(* IEC 61131-3 sources: PLC-IsaVODE/PLC-IsaVODE/samples/plc-programs (part 15) *)

(* ---- 331-SCALE_B2.ST ---- *)
FUNCTION _BYTE_TO_REAL:REAL
	VAR_INPUT
		IN :	BYTE;
	END_VAR

	_BYTE_TO_REAL := USINT_TO_REAL(BYTE_TO_USINT(IN));
END_FUNCTION

FUNCTION SCALE_B2:REAL
	VAR_INPUT
		IN1 :	BYTE;
		IN2 :	BYTE;
		K :	REAL;
		O :	REAL;
		IN1_MIN :	REAL;
		IN1_MAX :	REAL;
		IN2_MIN :	REAL;
		IN2_MAX :	REAL;
	END_VAR

	SCALE_B2 := 	(((in1_max - in1_min)* _BYTE_TO_REAL(in1) + (in2_max - in2_min)* _BYTE_TO_REAL(in2)) * 0.003921569 + in1_min + in2_min) * K + O;

END_FUNCTION

PROGRAM program0
  VAR
	IN1 :	BYTE;
	IN2 :	BYTE;
	K :	REAL;
	O :	REAL;
	IN1_MIN :	REAL;
	IN1_MAX :	REAL;
	IN2_MIN :	REAL;
	IN2_MAX :	REAL;
	CEIL5_OUT : REAL;
  END_VAR

  CEIL5_OUT := SCALE_B2(IN1, IN2, K, O, IN1_MIN, IN1_MAX, IN2_MIN, IN2_MAX);

END_PROGRAM

CONFIGURATION Config0

  RESOURCE Res0 ON PLC
    TASK task0(INTERVAL := T#20ms,PRIORITY := 0);
    PROGRAM instance0 WITH task0 : program0;
  END_RESOURCE
END_CONFIGURATION

(* ---- 334-AIR_ENTHALPY.ST ---- *)
FUNCTION SDD:REAL

	VAR_INPUT
		T :	REAL;
		ICE :	BOOL;
	END_VAR

	IF ice THEN
		SDD := 611.153 * EXP(22.4433 * T / (272.186 + T));
	ELSE
		SDD := 611.213 * EXP(17.5043 * T / (241.2 + T));
	END_IF;

END_FUNCTION

FUNCTION DEW_CON:REAL

	VAR_INPUT
		RH :	REAL;
		T :	REAL;
	END_VAR

	IF RH > 0.0 AND T > -50.0 THEN
		DEW_CON := 2.166824303E-2 * RH * SDD(T,FALSE)  / (T - -273.15);
	ELSE
		DEW_CON := 0.0;
	END_IF;

END_FUNCTION

FUNCTION AIR_ENTHALPY:REAL

	VAR_INPUT
		T :	REAL;
		RH :	REAL;
	END_VAR

	Air_enthalpy := 1.00482 * T + (1.86 * T + 2500.78) * dew_con(RH,T);

END_FUNCTION

PROGRAM program0
  VAR
    T :	REAL;
	RH :	REAL;
    CEIL5_OUT : REAL;
  END_VAR

  CEIL5_OUT := AIR_ENTHALPY(T, RH);
END_PROGRAM

CONFIGURATION Config0

  RESOURCE Res0 ON PLC
    TASK task0(INTERVAL := T#20ms,PRIORITY := 0);
    PROGRAM instance0 WITH task0 : program0;
  END_RESOURCE
END_CONFIGURATION

(* ---- 335-FRMP_B.ST ---- *)
FUNCTION FRMP_B:BYTE

	VAR_INPUT
		START :	BYTE;
		DIR :	BOOL;
		TD :	TIME;
		TR :	TIME;
	END_VAR

	IF TD < TR THEN
		FRMP_B := MIN(UDINT_TO_BYTE(DWORD_TO_UDINT(SHL(TIME_TO_DWORD(TD), 8)) / TIME_TO_UDINT(TR)), SEL(DIR, START, USINT_TO_BYTE(USINT#255 - BYTE_TO_USINT(START))));
		IF DIR THEN
			FRMP_B := USINT_TO_BYTE(BYTE_TO_USINT(START) + BYTE_TO_USINT(FRMP_B));
		ELSE
			FRMP_B := USINT_TO_BYTE(BYTE_TO_USINT(START) - BYTE_TO_USINT(FRMP_B));
		END_IF;
	ELSE
		FRMP_B := SEL(DIR, BYTE#0, BYTE#255);
	END_IF;
END_FUNCTION

PROGRAM program0
  VAR
    LocalVar0 : BYTE;
	LocalVar1 : BOOL;
	LocalVar2 : TIME;
	LocalVar3 : TIME;
    LocalOUT  : BYTE;
  END_VAR

  LocalOUT := FRMP_B(LocalVar0, LocalVar1, LocalVar2,LocalVar3);
END_PROGRAM

CONFIGURATION Config0
  RESOURCE Res0 ON PLC
    TASK task0(INTERVAL := T#20ms,PRIORITY := 0);
    PROGRAM instance0 WITH task0 : program0;
  END_RESOURCE
END_CONFIGURATION

(* ---- 336-MD5_AUX.ST ---- *)
FUNCTION MD5_AUX:DWORD

	VAR_INPUT
		N :	INT;
		A :	DWORD;
		B :	DWORD;
		C :	DWORD;
		D :	DWORD;
		X :	DWORD;
		U :	INT;
		T :	DWORD;
	END_VAR

	VAR
		w :	DWORD;
	END_VAR

	CASE N OF
		1: w := (B AND C) OR (NOT(B) AND D);
		2: w := (B AND D) OR (C AND NOT D);
		3: w := (B XOR C XOR D);
		4: w := (C XOR (B OR  NOT(D)));
	END_CASE;

	MD5_AUX := UDINT_TO_DWORD(DWORD_TO_UDINT(B) + DWORD_TO_UDINT(ROL_DWORD(UDINT_TO_DWORD(DWORD_TO_UDINT(A) + DWORD_TO_UDINT(w) + DWORD_TO_UDINT(X) + DWORD_TO_UDINT(T)),U)));

END_FUNCTION

PROGRAM program0
	VAR
		N :	INT;
		A :	DWORD;
		B :	DWORD;
		C :	DWORD;
		D :	DWORD;
		X :	DWORD;
		U :	INT;
		T :	DWORD;
		CEIL5_OUT : DWORD;
	END_VAR

  	CEIL5_OUT := MD5_AUX(N, A, B, C, D, X, U, T);
END_PROGRAM

CONFIGURATION Config0

  RESOURCE Res0 ON PLC
    TASK task0(INTERVAL := T#20ms,PRIORITY := 0);
    PROGRAM instance0 WITH task0 : program0;
  END_RESOURCE
END_CONFIGURATION

(* ---- 34-TIME_TO_INT.ST ---- *)
FUNCTION TIME_TO_INT1:INT

VAR_INPUT
	IN :	TIME;
END_VAR

TIME_TO_INT1 := DINT_TO_INT(TIME_TO_DINT(IN));
END_FUNCTION

PROGRAM program0
  VAR
	IN :	TIME;
    CEIL5_OUT : INT;
  END_VAR

  CEIL5_OUT := TIME_TO_INT1(IN);
END_PROGRAM

CONFIGURATION Config0

  RESOURCE Res0 ON PLC
    TASK task0(INTERVAL := T#20ms,PRIORITY := 0);
    PROGRAM instance0 WITH task0 : program0;
  END_RESOURCE
END_CONFIGURATION

(* ---- 35-C_TO_F.ST ---- *)
FUNCTION C_TO_F:REAL
	VAR_INPUT
		CELSIUS :	REAL;
	END_VAR

	C_TO_F := celsius * 1.8 + 32.0;
END_FUNCTION

PROGRAM program0
  VAR
    LocalVar0 : REAL;
    CEIL5_OUT : REAL;
  END_VAR

  CEIL5_OUT := C_TO_F(LocalVar0);
END_PROGRAM

CONFIGURATION Config0

  RESOURCE Res0 ON PLC
    TASK task0(INTERVAL := T#20ms,PRIORITY := 0);
    PROGRAM instance0 WITH task0 : program0;
  END_RESOURCE
END_CONFIGURATION

(* ---- 355-MULTIME.ST ---- *)
FUNCTION _REAL_TO_DWORD: DWORD

  VAR_INPUT
    X :	REAL;
  END_VAR

  IF REAL_TO_DWORD(0.5) = DWORD#1 THEN
    _REAL_TO_DWORD := REAL_TO_DWORD(x);
  ELSIF X > 0.0 THEN
    _REAL_TO_DWORD := REAL_TO_DWORD(x+0.5);
  ELSIF X < 0.0 THEN
    _REAL_TO_DWORD := REAL_TO_DWORD(x-0.5);
  ELSE
    _REAL_TO_DWORD := DWORD#0;
  END_IF;
END_FUNCTION

FUNCTION _DWORD_TO_REAL:REAL
	VAR_INPUT
		IN :	DWORD;
	END_VAR

	_DWORD_TO_REAL := UDINT_TO_REAL(DWORD_TO_UDINT(IN));

END_FUNCTION

FUNCTION MULTIME:TIME
	VAR_INPUT
		T :	TIME;
		M :	REAL;
	END_VAR

	multime := DWORD_TO_TIME(_REAL_TO_DWORD(_DWORD_TO_REAL(TIME_TO_DWORD(t))*M));
END_FUNCTION

PROGRAM program0
  VAR
    LocalVar0 : TIME;
	LocalVar1 : REAL;
	LocalOUT  : TIME;
  END_VAR
  	LocalOUT := MULTIME(LocalVar0, LocalVar1);
END_PROGRAM

CONFIGURATION Config0
  RESOURCE Res0 ON PLC
    TASK task0(INTERVAL := T#20ms,PRIORITY := 0);
    PROGRAM instance0 WITH task0 : program0;
  END_RESOURCE
END_CONFIGURATION

(* ---- 356-OFFSET2.ST ---- *)
FUNCTION OFFSET2:REAL

	VAR_INPUT
		X :	REAL;
		O1 :	BOOL;
		O2 :	BOOL;
		O3 :	BOOL;
		O4 :	BOOL;
		D :	BOOL;
		OFFSET_1 :	REAL;
		OFFSET_2 :	REAL;
		OFFSET_3 :	REAL;
		OFFSET_4 :	REAL;
		DEFAULT :	REAL;
	END_VAR

	IF D THEN Offset2 := default; ELSE Offset2 := X; END_IF;
	IF O4 THEN Offset2 := Offset2 + offset_4;
	ELSIF O3 THEN Offset2 := Offset2 + offset_3;
	ELSIF O2 THEN Offset2 := Offset2 + offset_2;
	ELSIF O1 THEN Offset2 := Offset2 + offset_1;
	END_IF;

END_FUNCTION

PROGRAM program0
	VAR
		X :	REAL;
		O1 :	BOOL;
		O2 :	BOOL;
		O3 :	BOOL;
		O4 :	BOOL;
		D :	BOOL;
		OFFSET_1 :	REAL;
		OFFSET_2 :	REAL;
		OFFSET_3 :	REAL;
		OFFSET_4 :	REAL;
		DEFAULT :	REAL;
		OUT : REAL;
	END_VAR

	OUT := OFFSET2(X, O1, O2, O3, O4, D, OFFSET_1, OFFSET_2, OFFSET_3, OFFSET_4, DEFAULT);
END_PROGRAM

CONFIGURATION Config0

	RESOURCE Res0 ON PLC
		TASK task0(INTERVAL := T#20ms,PRIORITY := 0);
		PROGRAM instance0 WITH task0 : program0;
	END_RESOURCE

END_CONFIGURATION

(* ---- 36-DATE_TO_UDINT.ST ---- *)
FUNCTION DATE_TO_UDINT2:UDINT
	VAR_INPUT
		IN :	UDINT;
	END_VAR

	DATE_TO_UDINT2 := IN;
END_FUNCTION

PROGRAM program0
  VAR
    LocalVar0 : UDINT;
	LocalOUT  : UDINT;
  END_VAR
  	LocalOUT := DATE_TO_UDINT2(LocalVar0);
END_PROGRAM

CONFIGURATION Config0
  RESOURCE Res0 ON PLC
    TASK task0(INTERVAL := T#20ms,PRIORITY := 0);
    PROGRAM instance0 WITH task0 : program0;
  END_RESOURCE
END_CONFIGURATION

(* ---- 363-OFFSET.ST ---- *)
FUNCTION _OFFSET:REAL

	VAR_INPUT
		X :	REAL;
		O1 :	BOOL;
		O2 :	BOOL;
		O3 :	BOOL;
		O4 :	BOOL;
		D :	BOOL;
		OFFSET_1 :	REAL;
		OFFSET_2 :	REAL;
		OFFSET_3 :	REAL;
		OFFSET_4 :	REAL;
		DEFAULT :	REAL;
	END_VAR

	IF D THEN _Offset := default; ELSE _Offset := X; END_IF;
	IF O1 THEN _Offset := _Offset + offset_1; END_IF;
	IF O2 THEN _Offset := _Offset + offset_2; END_IF;
	IF O3 THEN _Offset := _Offset + offset_3; END_IF;
	IF O4 THEN _Offset := _Offset + offset_4; END_IF;

END_FUNCTION

PROGRAM program0

	VAR
		X :	REAL;
		O1 :	BOOL;
		O2 :	BOOL;
		O3 :	BOOL;
		O4 :	BOOL;
		D :	BOOL;
		OFFSET_1 :	REAL;
		OFFSET_2 :	REAL;
		OFFSET_3 :	REAL;
		OFFSET_4 :	REAL;
		DEFAULT :	REAL;
		OUT : REAL;
	END_VAR

	OUT := _OFFSET(X, O1, O2, O3, O4, D, OFFSET_1, OFFSET_2, OFFSET_3, OFFSET_4, DEFAULT);
END_PROGRAM

CONFIGURATION Config0

	RESOURCE Res0 ON PLC
		TASK task0(INTERVAL := T#20ms,PRIORITY := 0);
		PROGRAM instance0 WITH task0 : program0;
	END_RESOURCE

END_CONFIGURATION

(* ---- 365-CMP.ST ---- *)
FUNCTION EXP10 : REAL
  VAR_INPUT
    x : REAL;
  END_VAR

  exp10 := EXP(X * 2.30258509299405);
  (* from OSCAT library; www.oscat.de  *)
END_FUNCTION

FUNCTION FLOOR : INT
  VAR_INPUT
    x : REAL;
  END_VAR

  FLOOR := REAL_TO_INT(X);
  IF INT_TO_REAL(FLOOR) > X THEN
  	floor := floor - 1;
  END_IF;
  (* from OSCAT library; www.oscat.de  *)
END_FUNCTION

FUNCTION CMP:BOOL
	VAR_INPUT
		X :	REAL;
		Y :	REAL;
		N :	INT;
	END_VAR

	VAR
		tmp :	REAL;
	END_VAR

	tmp := ABS(x);
	IF tmp > 0.0 THEN
		tmp := EXP10(INT_TO_REAL(FLOOR(LOG(tmp))-N+1));
	ELSE
		tmp := EXP10(tmp);
	END_IF;
	CMP := ABS(X - Y) < tmp;

END_FUNCTION

PROGRAM program0
  VAR
    LocalVar0 : REAL;
    LocalVar1 : REAL;
	LocalVar2 : INT;
    CEIL5_OUT : BOOL;
  END_VAR

  CEIL5_OUT := CMP(LocalVar0, LocalVar1, LocalVar2);
END_PROGRAM

CONFIGURATION Config0

  RESOURCE Res0 ON PLC
    TASK task0(INTERVAL := T#20ms,PRIORITY := 0);
    PROGRAM instance0 WITH task0 : program0;
  END_RESOURCE
END_CONFIGURATION

(* ---- 37-LEAP_DAY.ST ---- *)
FUNCTION LEAP_DAY:BOOL

	VAR_INPUT
		IDATE :	UDINT;
	END_VAR

	LEAP_DAY := IDATE MOD UDINT#126230400 = UDINT#68169600;

END_FUNCTION

PROGRAM program0
	VAR
		IDATE :	UDINT;
		OUT : BOOL;
	END_VAR

	OUT := LEAP_DAY(IDATE);
END_PROGRAM

CONFIGURATION Config0

	RESOURCE Res0 ON PLC
		TASK task0(INTERVAL := T#20ms,PRIORITY := 0);
		PROGRAM instance0 WITH task0 : program0;
	END_RESOURCE

END_CONFIGURATION

(* ---- 370-SET_TOD.ST ---- *)
FUNCTION _REAL_TO_UDINT:UDINT

	VAR_INPUT
		X :	REAL;
	END_VAR

	IF REAL_TO_UDINT(0.5) = UDINT#1 THEN
		_REAL_TO_UDINT := REAL_TO_UDINT(x);
	ELSIF X > 0.0 THEN
		_REAL_TO_UDINT := REAL_TO_UDINT(x+0.5);
	ELSIF X < 0.0 THEN
		_REAL_TO_UDINT := REAL_TO_UDINT(x-0.5);
	ELSE
		_REAL_TO_UDINT := UDINT#0;
	END_IF;

END_FUNCTION

FUNCTION _INT_TO_UDINT:UDINT

	VAR_INPUT
		IN :	INT;
	END_VAR

	_INT_TO_UDINT := DINT_TO_UDINT(INT_TO_DINT(IN));

END_FUNCTION

FUNCTION SET_TOD:UDINT

	VAR_INPUT
		HOUR :	INT;
		MINUTE :	INT;
		SECOND :	REAL;
	END_VAR

	set_Tod := _REAL_TO_UDINT(second * 1000.0) + _INT_TO_UDINT(minute) * UDINT#60000 + _INT_TO_UDINT(hour) * UDINT#3600000;

END_FUNCTION

PROGRAM program0

	VAR
		HOUR :	INT;
		MINUTE :	INT;
		SECOND :	REAL;
		CEIL5_OUT : UDINT;
	END_VAR

	CEIL5_OUT := SET_TOD(HOUR, MINUTE, SECOND);

END_PROGRAM

CONFIGURATION Config0

	RESOURCE Res0 ON PLC
		TASK task0(INTERVAL := T#20ms,PRIORITY := 0);
		PROGRAM instance0 WITH task0 : program0;
	END_RESOURCE

END_CONFIGURATION

(* ---- 371-HEAT_INDEX.ST ---- *)
FUNCTION C_TO_F:REAL
	VAR_INPUT
		CELSIUS :	REAL;
	END_VAR

	C_TO_F := celsius * 1.8 + 32.0;
END_FUNCTION

FUNCTION F_TO_C:REAL
	VAR_INPUT
		FAHRENHEIT :	REAL;
	END_VAR
	F_TO_C := (fahrenheit - 32.0) * 0.5555555555555;
END_FUNCTION

FUNCTION HEAT_INDEX:REAL

	VAR_INPUT
		T :	REAL;
		RH :	REAL;
	END_VAR

	VAR
		RH2 :	REAL;
		T2 :	REAL;
		TX :	REAL;
	END_VAR

	IF RH < 20.0 OR T < 20.0 THEN
		HEAT_INDEX := T;
	ELSE
		TX := T;
		RH2 := RH * RH;
		TX := C_TO_F(TX);
		T2 := TX * TX;
		HEAT_INDEX := -42.379 + 2.04901523 * TX - 6.83783E-3 * T2
				+ RH * (10.1433127 - 0.22475541 * TX + 1.22874E-3 * T2)
				+ RH2 * (8.5282E-4 * TX - 5.481717E-2 - 1.99E-6 * T2);
		HEAT_INDEX := F_TO_C(HEAT_INDEX);
	END_IF;

END_FUNCTION

PROGRAM program0
  VAR
    T :	REAL;
	RH :	REAL;
    CEIL5_OUT : REAL;
  END_VAR

  CEIL5_OUT := HEAT_INDEX(T, RH);
END_PROGRAM

CONFIGURATION Config0

  RESOURCE Res0 ON PLC
    TASK task0(INTERVAL := T#20ms,PRIORITY := 0);
    PROGRAM instance0 WITH task0 : program0;
  END_RESOURCE
END_CONFIGURATION

(* ---- 38-TOD_TO_TIME.ST ---- *)
FUNCTION TOD_TO_TIME:TIME
	VAR_INPUT
		IN :	UDINT;
	END_VAR

	TOD_TO_TIME := DWORD_TO_TIME(UDINT_TO_DWORD(IN));
END_FUNCTION

PROGRAM program0
  VAR
	IN :	UDINT;
    CEIL5_OUT : TIME;
  END_VAR

  CEIL5_OUT := TOD_TO_TIME(IN);
END_PROGRAM

CONFIGURATION Config0

  RESOURCE Res0 ON PLC
    TASK task0(INTERVAL := T#20ms,PRIORITY := 0);
    PROGRAM instance0 WITH task0 : program0;
  END_RESOURCE
END_CONFIGURATION

(* ---- 384-EXPN.ST ---- *)
FUNCTION BIT_OF_DWORD : BOOL
  VAR_INPUT
    IN : DWORD;
    N : INT;
  END_VAR

  BIT_OF_DWORD := (SHR(in,N) AND 16#00000001) > 0;
END_FUNCTION

FUNCTION EXPN:REAL

	VAR_INPUT
		X :	REAL;
		N :	INT;
	END_VAR

	VAR
		N_word :	WORD;
		X_tmp :	REAL;
		sign :	BOOL;
	END_VAR

	N_word := INT_TO_WORD(N);
	X_tmp := X;
	sign := BIT_OF_DWORD(WORD_TO_DWORD(N_word),15);
	N_word := INT_TO_WORD(ABS(N));
	IF BIT_OF_DWORD(WORD_TO_DWORD(N_word),0) THEN expn := X_tmp; ELSE expn := 1.0; END_IF;    (* N_word.X0 *)
	N_word := SHR(N_word,1);
	WHILE N_word > WORD#0 DO
		X_tmp := X_tmp * X_tmp;
		IF BIT_OF_DWORD(WORD_TO_DWORD(N_word),0) THEN expn := expn * X_tmp; END_IF;       (* N_word.X0 *)
		N_word := SHR(N_word,1);
	END_WHILE;
	IF sign THEN EXPN := 1.0 / EXPN; END_IF;

END_FUNCTION

PROGRAM program0
  VAR
    LocalVar0 : REAL;
	LocalVar1 : INT;
	LocalOUT  : REAL;
  END_VAR
  	LocalOUT := EXPN(LocalVar0, LocalVar1);
END_PROGRAM

CONFIGURATION Config0
  RESOURCE Res0 ON PLC
    TASK task0(INTERVAL := T#20ms,PRIORITY := 0);
    PROGRAM instance0 WITH task0 : program0;
  END_RESOURCE
END_CONFIGURATION

(* ---- 385-ROUND.ST ---- *)
FUNCTION _REAL_TO_DINT:DINT
	VAR_INPUT
		X :	REAL;
	END_VAR

	IF REAL_TO_DINT(0.5) = DINT#1 THEN
		_REAL_TO_DINT := REAL_TO_DINT(x);
		RETURN;
	END_IF;

	IF X > 0.0 THEN
		_REAL_TO_DINT := REAL_TO_DINT(x+0.5);
	ELSIF X < 0.0 THEN
		_REAL_TO_DINT := REAL_TO_DINT(x-0.5);
	ELSE
		_REAL_TO_DINT := DINT#0;
	END_IF;
END_FUNCTION

FUNCTION ROUND:REAL

	VAR_INPUT
		IN :	REAL;
		N :	INT;
	END_VAR

	VAR
		X :	REAL;
	END_VAR

	IF N < 4 THEN
		IF N < 2 THEN
			IF N = 0 THEN X := 1.0; ELSE X := 10.0; END_IF;
		ELSE
			IF N = 2 THEN X := 100.0; ELSE X := 1000.0; END_IF;
		END_IF;
	ELSE
		IF N < 6 THEN
			IF N = 4 THEN X := 10000.0; ELSE X := 100000.0; END_IF;
		ELSE
			IF N = 6 THEN X := 1000000.0; ELSE X := 10000000.0; END_IF;
		END_IF;
	END_IF;

	ROUND := DINT_TO_REAL(_REAL_TO_DINT(in * X)) / X;

END_FUNCTION

PROGRAM program0
	VAR
		IN : REAL;
		N :	INT;
		X :	REAL;
	END_VAR
		X := ROUND(IN, N);
END_PROGRAM

CONFIGURATION Config0

	RESOURCE Res0 ON PLC
		TASK task0(INTERVAL := T#20ms,PRIORITY := 0);
		PROGRAM instance0 WITH task0 : program0;
	END_RESOURCE

END_CONFIGURATION

(* ---- 39-DATE_TO_REAL.ST ---- *)
FUNCTION DATE_TO_REAL2:REAL
	VAR_INPUT
		IN :	UDINT;
	END_VAR

	DATE_TO_REAL2 := UDINT_TO_REAL(IN);
END_FUNCTION

PROGRAM program0
  VAR
    LocalVar0 : UDINT;
	LocalOUT  : REAL;
  END_VAR
  	LocalOUT := DATE_TO_REAL2(LocalVar0);
END_PROGRAM

CONFIGURATION Config0
  RESOURCE Res0 ON PLC
    TASK task0(INTERVAL := T#20ms,PRIORITY := 0);
    PROGRAM instance0 WITH task0 : program0;
  END_RESOURCE
END_CONFIGURATION

(* ---- 395-SET_DATE.ST ---- *)
FUNCTION _INT_TO_UDINT:UDINT
	VAR_INPUT
		IN :	INT;
	END_VAR

	_INT_TO_UDINT := DINT_TO_UDINT(INT_TO_DINT(IN));
END_FUNCTION

FUNCTION SET_DATE:UDINT

	VAR_INPUT
		YEAR :	INT;
		MONTH :	INT;
		DAY :	INT;
	END_VAR

	VAR
		count :	INT;
	END_VAR

	IF month > 2 THEN
		count := (month - 1) * 30;
		IF month > 7 THEN
			count := count + DWORD_TO_INT(SHR(DINT_TO_DWORD(INT_TO_DINT(month) - INT_TO_DINT(3)),1));
		ELSE
			count := count + DWORD_TO_INT(SHR(DINT_TO_DWORD(INT_TO_DINT(month) - INT_TO_DINT(4)),1));
		END_IF;
		IF SHL(INT_TO_WORD(year),14) = WORD#0 THEN
			count := count + 1;
		END_IF;
	ELSE
		count := (month - 1) * 31;
	END_IF;
	SET_DATE := (_INT_TO_UDINT(count + day - 1) + DWORD_TO_UDINT(SHR(UDINT_TO_DWORD(_INT_TO_UDINT(year) * UDINT#1461 - UDINT#2878169), 2))) * UDINT#86400;

END_FUNCTION

PROGRAM program0
  VAR
	YEAR :	INT;
	MONTH :	INT;
	DAY :	INT;
    CEIL5_OUT : UDINT;
  END_VAR

  CEIL5_OUT := SET_DATE(YEAR, MONTH, DAY);
END_PROGRAM

CONFIGURATION Config0

  RESOURCE Res0 ON PLC
    TASK task0(INTERVAL := T#20ms,PRIORITY := 0);
    PROGRAM instance0 WITH task0 : program0;
  END_RESOURCE
END_CONFIGURATION

(* ---- 40-DWORD_TO_DT.ST ---- *)
FUNCTION DWORD_TO_DT2:UDINT

	VAR_INPUT
		IN :	DWORD;
	END_VAR

	DWORD_TO_DT2 := DWORD_TO_UDINT(IN);
END_FUNCTION

PROGRAM program0
  VAR
    LocalVar0 : DWORD;
	LocalOUT  : UDINT;
  END_VAR
  	LocalOUT := DWORD_TO_DT2(LocalVar0);
END_PROGRAM

CONFIGURATION Config0
  RESOURCE Res0 ON PLC
    TASK task0(INTERVAL := T#20ms,PRIORITY := 0);
    PROGRAM instance0 WITH task0 : program0;
  END_RESOURCE
END_CONFIGURATION

(* ---- 400-TEMP_PT.ST ---- *)
FUNCTION RES_PT:REAL
	VAR_INPUT
		T :	REAL;
		R0 :	REAL;
	END_VAR

	VAR
		T2 :	REAL;
	END_VAR

	T2 := T * T;

	IF T >= 0.0 THEN
		RES_PT := R0 * ( 1.0 + 3.90802E-3 * T + -5.802E-7 * T2);
	ELSE
		RES_PT := R0 * ( 1.0 + 3.90802E-3 * T + -5.802E-7 * T2 + -4.27350E-12 * (T - 100.0) * T2 * T);
	END_IF;

END_FUNCTION

FUNCTION TEMP_PT:REAL

	VAR_INPUT
		RES :	REAL;
		R0 :	REAL;
	END_VAR

	VAR
		step_var :	REAL := REAL#50.0;
		X :	REAL;
		Y :	REAL;
		t1 :	REAL;
	END_VAR

	X := 3.9083E-3 * R0;
	Y := -5.775E-7 * R0;
	IF Res >= R0 THEN
		t1 := X * X - 4.0 * Y * (R0 - Res);
		IF t1 < 0.0 THEN
			TEMP_PT := 10000.0;
		ELSE
			TEMP_PT := (-X + SQRT(t1)) / (2.0 * Y);
		END_IF;
	ELSE
		TEMP_PT := -100.0;
		WHILE step_var > 0.01 DO
			IF RES_PT(TEMP_PT, R0) < res THEN TEMP_PT := TEMP_PT + step_var; ELSE TEMP_PT := TEMP_PT - step_var; END_IF;
			step_var := step_var * 0.5;
		END_WHILE;
	END_IF;
END_FUNCTION

PROGRAM program0
	VAR
		RES :	REAL;
		R0 :	REAL;
		CEIL5_OUT : REAL;
	END_VAR

	CEIL5_OUT := TEMP_PT(RES, R0);
END_PROGRAM

CONFIGURATION Config0
	RESOURCE Res0 ON PLC
		TASK task0(INTERVAL := T#20ms,PRIORITY := 0);
		PROGRAM instance0 WITH task0 : program0;
	END_RESOURCE
END_CONFIGURATION

(* ---- 404-MONTH_OF_DATE.ST ---- *)
FUNCTION LEAP_OF_DATE:BOOL

	VAR_INPUT
		IDATE :	UDINT;
	END_VAR

	LEAP_OF_DATE := SHL(UDINT_TO_DWORD((idate + UDINT#43200) / UDINT#31557600), 30) = DWORD#16#80000000;

END_FUNCTION

FUNCTION DAY_OF_YEAR:INT
	VAR_INPUT
		IDATE :	DATE;
	END_VAR

	DAY_OF_YEAR := UDINT_TO_INT((DATE_TO_UDINT(idate) / UDINT#86400) MOD UDINT#1461);
	IF DAY_OF_YEAR > 729 THEN
		IF DAY_OF_YEAR > 1095 THEN DAY_OF_YEAR := DAY_OF_YEAR - 1095; ELSE DAY_OF_YEAR := DAY_OF_YEAR - 729; END_IF;
	ELSIF DAY_OF_YEAR > 364 THEN
		DAY_OF_YEAR := DAY_OF_YEAR - 364;
	ELSE
		DAY_OF_YEAR := DAY_OF_YEAR + 1;
	END_IF;
END_FUNCTION

FUNCTION MONTH_OF_DATE:INT

	VAR_INPUT
		IDATE :	DATE;
	END_VAR

	MONTH_OF_DATE := DAY_OF_YEAR(idate);
	IF MONTH_OF_DATE < 32 THEN
		MONTH_OF_DATE := 1;
	ELSIF LEAP_OF_DATE(DATE_TO_UDINT(IDATE)) THEN
		MONTH_OF_DATE := (MONTH_OF_DATE * 53 + 1668) / 1623;
	ELSE
		MONTH_OF_DATE := (MONTH_OF_DATE * 53 + 1700) / 1620;
	END_IF;

END_FUNCTION

PROGRAM program0
  VAR
    LocalVar0 : DATE;
	LocalOUT  : INT;
  END_VAR
  	LocalOUT := MONTH_OF_DATE(LocalVar0);
END_PROGRAM

CONFIGURATION Config0
  RESOURCE Res0 ON PLC
    TASK task0(INTERVAL := T#20ms,PRIORITY := 0);
    PROGRAM instance0 WITH task0 : program0;
  END_RESOURCE
END_CONFIGURATION

(* ---- 405-SCALE_B4.ST ---- *)
FUNCTION _BYTE_TO_REAL:REAL
	VAR_INPUT
		IN :	BYTE;
	END_VAR

	_BYTE_TO_REAL := USINT_TO_REAL(BYTE_TO_USINT(IN));
END_FUNCTION

FUNCTION SCALE_B4:REAL

	VAR_INPUT
		IN1 :	BYTE;
		IN2 :	BYTE;
		IN3 :	BYTE;
		IN4 :	BYTE;
		K :	REAL;
		O :	REAL;
		IN1_MIN :	REAL;
		IN1_MAX :	REAL;
		IN2_MIN :	REAL;
		IN2_MAX :	REAL;
		IN3_MIN :	REAL;
		IN3_MAX :	REAL;
		IN4_MIN :	REAL;
		IN4_MAX :	REAL;
	END_VAR

	SCALE_B4 := 	(((in1_max - in1_min)* _BYTE_TO_REAL(in1) + (in2_max - in2_min)* _BYTE_TO_REAL(in2) + (in3_max - in3_min)* _BYTE_TO_REAL(in3) + (in4_max - in4_min)* _BYTE_TO_REAL(in4))* 0.003921569 + in1_min + in2_min + in3_min + in4_min) * K + O;

END_FUNCTION

PROGRAM program0
  VAR
	IN1 :	BYTE;
	IN2 :	BYTE;
	IN3 :	BYTE;
	IN4 :	BYTE;
	K :	REAL;
	O :	REAL;
	IN1_MIN :	REAL;
	IN1_MAX :	REAL;
	IN2_MIN :	REAL;
	IN2_MAX :	REAL;
	IN3_MIN :	REAL;
	IN3_MAX :	REAL;
	IN4_MIN :	REAL;
	IN4_MAX :	REAL;
	CEIL5_OUT : REAL;
  END_VAR

  CEIL5_OUT := SCALE_B4(IN1, IN2, IN3, IN4, K, O, IN1_MIN, IN1_MAX, IN2_MIN, IN2_MAX, IN3_MIN, IN3_MAX, IN4_MIN, IN4_MAX);

END_PROGRAM

CONFIGURATION Config0

  RESOURCE Res0 ON PLC
    TASK task0(INTERVAL := T#20ms,PRIORITY := 0);
    PROGRAM instance0 WITH task0 : program0;
  END_RESOURCE
END_CONFIGURATION

(* ---- 408-SCALE_X4.ST ---- *)
FUNCTION SCALE_X4:REAL
	VAR_INPUT
		IN1 :	BOOL;
		IN2 :	BOOL;
		IN3 :	BOOL;
		IN4 :	BOOL;
		K :	REAL;
		O :	REAL;
		IN1_MIN :	REAL;
		IN1_MAX :	REAL;
		IN2_MIN :	REAL;
		IN2_MAX :	REAL;
		IN3_MIN :	REAL;
		IN3_MAX :	REAL;
		IN4_MIN :	REAL;
		IN4_MAX :	REAL;
	END_VAR
	IF NOT in1 THEN scale_X4 := in1_min; ELSE scale_X4 := in1_max; END_IF;
	IF NOT in2 THEN scale_x4 := scale_x4 + in2_min; ELSE scale_x4 := scale_x4 + in2_max; END_IF;
	IF NOT in3 THEN scale_x4 := scale_x4 + in3_min; ELSE scale_x4 := scale_x4 + in3_max; END_IF;
	IF NOT in4 THEN scale_x4 := scale_x4 + in4_min; ELSE scale_x4 := scale_x4 + in4_max; END_IF;
	scale_X4 := scale_X4 * k + O;
	END_FUNCTION

PROGRAM program0

  	VAR
		IN1 :	BOOL;
		IN2 :	BOOL;
		IN3 :	BOOL;
		IN4 :	BOOL;
		K :	REAL;
		O :	REAL;
		IN1_MIN :	REAL;
		IN1_MAX :	REAL;
		IN2_MIN :	REAL;
		IN2_MAX :	REAL;
		IN3_MIN :	REAL;
		IN3_MAX :	REAL;
		IN4_MIN :	REAL;
		IN4_MAX :	REAL;
		CEIL5_OUT : REAL;
  	END_VAR

  	CEIL5_OUT := SCALE_X4(IN1, IN2, IN3, IN4, K, O, IN1_MIN, IN1_MAX, IN2_MIN, IN2_MAX, IN3_MIN, IN3_MAX, IN4_MIN, IN4_MAX);
END_PROGRAM

CONFIGURATION Config0

	RESOURCE Res0 ON PLC
		TASK task0(INTERVAL := T#20ms,PRIORITY := 0);
		PROGRAM instance0 WITH task0 : program0;
	END_RESOURCE

END_CONFIGURATION

(* ---- 41-BYTE_TO_GRAY.ST ---- *)
FUNCTION BYTE_TO_GRAY:BYTE
	VAR_INPUT
		IN :	BYTE;
	END_VAR

	BYTE_TO_GRAY := IN XOR SHR(IN,1);
END_FUNCTION

PROGRAM program0
  VAR
    LocalVar0 : BYTE;
    CEIL5_OUT : BYTE;
  END_VAR

  CEIL5_OUT := BYTE_TO_GRAY(LocalVar0);
END_PROGRAM

CONFIGURATION Config0

  RESOURCE Res0 ON PLC
    TASK task0(INTERVAL := T#20ms,PRIORITY := 0);
    PROGRAM instance0 WITH task0 : program0;
  END_RESOURCE
END_CONFIGURATION

(* ---- 413-OSCAT_VERSION.ST ---- *)
FUNCTION _INT_TO_UDINT:UDINT
	VAR_INPUT
		IN :	INT;
	END_VAR

	_INT_TO_UDINT := DINT_TO_UDINT(INT_TO_DINT(IN));
END_FUNCTION

FUNCTION SET_DATE:UDINT

	VAR_INPUT
		YEAR :	INT;
		MONTH :	INT;
		DAY :	INT;
	END_VAR

	VAR
		count :	INT;
	END_VAR

	IF month > 2 THEN
		count := (month - 1) * 30;
		IF month > 7 THEN
			count := count + DWORD_TO_INT(SHR(DINT_TO_DWORD(INT_TO_DINT(month) - INT_TO_DINT(3)),1));
		ELSE
			count := count + DWORD_TO_INT(SHR(DINT_TO_DWORD(INT_TO_DINT(month) - INT_TO_DINT(4)),1));
		END_IF;
		IF SHL(INT_TO_WORD(year),14) = WORD#0 THEN
			count := count + 1;
		END_IF;
	ELSE
		count := (month - 1) * 31;
	END_IF;
	SET_DATE := (_INT_TO_UDINT(count + day - 1) + DWORD_TO_UDINT(SHR(UDINT_TO_DWORD(_INT_TO_UDINT(year) * UDINT#1461 - UDINT#2878169), 2))) * UDINT#86400;

END_FUNCTION

FUNCTION OSCAT_VERSION:DWORD

	VAR_INPUT
		IN :	BOOL;
	END_VAR

	IF in THEN
		Oscat_version := UDINT_TO_DWORD(set_Date(2012,01,02));
	ELSE
		Oscat_version := DWORD#333;
	END_IF;

END_FUNCTION

PROGRAM program0
	VAR
		IN :	BOOL;
		OUT : DWORD;
	END_VAR

	OUT := OSCAT_VERSION(IN);
END_PROGRAM

CONFIGURATION Config0

	RESOURCE Res0 ON PLC
		TASK task0(INTERVAL := T#20ms,PRIORITY := 0);
		PROGRAM instance0 WITH task0 : program0;
	END_RESOURCE

END_CONFIGURATION

(* ---- 417-NETWORK_VERSION.ST ---- *)
FUNCTION _INT_TO_UDINT:UDINT
	VAR_INPUT
		IN :	INT;
	END_VAR

	_INT_TO_UDINT := DINT_TO_UDINT(INT_TO_DINT(IN));
END_FUNCTION

FUNCTION SET_DATE:UDINT

	VAR_INPUT
		YEAR :	INT;
		MONTH :	INT;
		DAY :	INT;
	END_VAR

	VAR
		count :	INT;
	END_VAR

	IF month > 2 THEN
		count := (month - 1) * 30;
		IF month > 7 THEN
			count := count + DWORD_TO_INT(SHR(DINT_TO_DWORD(INT_TO_DINT(month) - INT_TO_DINT(3)),1));
		ELSE
			count := count + DWORD_TO_INT(SHR(DINT_TO_DWORD(INT_TO_DINT(month) - INT_TO_DINT(4)),1));
		END_IF;
		IF SHL(INT_TO_WORD(year),14) = WORD#0 THEN
			count := count + 1;
		END_IF;
	ELSE
		count := (month - 1) * 31;
	END_IF;
	SET_DATE := (_INT_TO_UDINT(count + day - 1) + DWORD_TO_UDINT(SHR(UDINT_TO_DWORD(_INT_TO_UDINT(year) * UDINT#1461 - UDINT#2878169), 2))) * UDINT#86400;

END_FUNCTION

FUNCTION NETWORK_VERSION:DWORD

	VAR_INPUT
		IN :	BOOL;
	END_VAR

	IF in THEN
		NETWORK_VERSION := UDINT_TO_DWORD(set_Date(2011,12,01));
	ELSE
		NETWORK_VERSION := DWORD#121;
	END_IF;

END_FUNCTION

PROGRAM program0
	VAR
		IN :	BOOL;
		CEIL5_OUT : DWORD;
	END_VAR

  	CEIL5_OUT := NETWORK_VERSION(IN);
END_PROGRAM

CONFIGURATION Config0

  RESOURCE Res0 ON PLC
    TASK task0(INTERVAL := T#20ms,PRIORITY := 0);
    PROGRAM instance0 WITH task0 : program0;
  END_RESOURCE
END_CONFIGURATION

(* ---- 419-BUILDING_VERSION.ST ---- *)
FUNCTION _INT_TO_UDINT:UDINT
	VAR_INPUT
		IN :	INT;
	END_VAR

	_INT_TO_UDINT := DINT_TO_UDINT(INT_TO_DINT(IN));
END_FUNCTION

FUNCTION SET_DATE:UDINT

	VAR_INPUT
		YEAR :	INT;
		MONTH :	INT;
		DAY :	INT;
	END_VAR

	VAR
		count :	INT;
	END_VAR

	IF month > 2 THEN
		count := (month - 1) * 30;
		IF month > 7 THEN
			count := count + DWORD_TO_INT(SHR(DINT_TO_DWORD(INT_TO_DINT(month) - INT_TO_DINT(3)),1));
		ELSE
			count := count + DWORD_TO_INT(SHR(DINT_TO_DWORD(INT_TO_DINT(month) - INT_TO_DINT(4)),1));
		END_IF;
		IF SHL(INT_TO_WORD(year),14) = WORD#0 THEN
			count := count + 1;
		END_IF;
	ELSE
		count := (month - 1) * 31;
	END_IF;
	SET_DATE := (_INT_TO_UDINT(count + day - 1) + DWORD_TO_UDINT(SHR(UDINT_TO_DWORD(_INT_TO_UDINT(year) * UDINT#1461 - UDINT#2878169), 2))) * UDINT#86400;

END_FUNCTION

FUNCTION BUILDING_VERSION:DWORD

	VAR_INPUT
		IN :	BOOL;
	END_VAR

	IF in THEN
		BUILDING_VERSION := UDINT_TO_DWORD(set_Date(2011,02,03));
	ELSE
		BUILDING_VERSION := DWORD#100;
	END_IF;

END_FUNCTION

PROGRAM program0
	VAR
		IN :	BOOL;
		CEIL5_OUT : DWORD;
	END_VAR

  	CEIL5_OUT := BUILDING_VERSION(IN);
END_PROGRAM

CONFIGURATION Config0

  RESOURCE Res0 ON PLC
    TASK task0(INTERVAL := T#20ms,PRIORITY := 0);
    PROGRAM instance0 WITH task0 : program0;
  END_RESOURCE
END_CONFIGURATION

(* ---- 42-F_TO_C.ST ---- *)
FUNCTION F_TO_C:REAL
	VAR_INPUT
		FAHRENHEIT :	REAL;
	END_VAR
	F_TO_C := (fahrenheit - 32.0) * 0.5555555555555;
END_FUNCTION

PROGRAM program0
  VAR
    LocalVar0 : REAL;
	LocalOUT  : REAL;
  END_VAR
  	LocalOUT := F_TO_C(LocalVar0);
END_PROGRAM

CONFIGURATION Config0
  RESOURCE Res0 ON PLC
    TASK task0(INTERVAL := T#20ms,PRIORITY := 0);
    PROGRAM instance0 WITH task0 : program0;
  END_RESOURCE
END_CONFIGURATION

(* ---- 421-GCD.ST ---- *)
FUNCTION GCD:INT

	VAR_INPUT
		A :	DINT;
		B :	DINT;
	END_VAR

	VAR
		t :	DINT;
		_A :	DINT;
		_B :	DINT;
	END_VAR

	_A := A;
	_B := B;

	IF _A = DINT#0 THEN
		GCD := DINT_TO_INT(ABS(_B));
	ELSIF _B = DINT#0 THEN
		GCD := DINT_TO_INT(ABS(_A));
	ELSE
		_A := ABS(_A);
		_B := ABS(_B);
		GCD := 1;

		WHILE NOT((DINT_TO_DWORD(_A) AND DWORD#1) > DWORD#0 OR (DINT_TO_DWORD(_B) AND DWORD#1) > DWORD#0) DO
			_A := DWORD_TO_DINT(SHR(DINT_TO_DWORD(_A),1));
			_B := DWORD_TO_DINT(SHR(DINT_TO_DWORD(_B),1));
			GCD := DWORD_TO_INT(SHR(INT_TO_DWORD(GCD),1));
		END_WHILE;
		WHILE _A > DINT#0 DO
			IF NOT((DINT_TO_DWORD(_A) AND DWORD#1) > DWORD#0) THEN
				_A := DWORD_TO_DINT(SHR(DINT_TO_DWORD(_A),1));
			ELSIF NOT((DINT_TO_DWORD(_B) AND DWORD#1) > DWORD#0) THEN
				_B := DWORD_TO_DINT(SHR(DINT_TO_DWORD(_B),1));
			ELSE
				t := DWORD_TO_DINT(SHR(DINT_TO_DWORD(ABS(_A-_B)),1));
				IF _A < _B THEN
					_B := t;
				ELSE
					_A := t;
				END_IF;
			END_IF;
		END_WHILE;
		GCD := GCD * DINT_TO_INT(_B);
	END_IF;

END_FUNCTION

PROGRAM program0
  VAR
    A :	DINT;
	B :	DINT;
    LocalOUT  : INT;
  END_VAR

  LocalOUT := GCD(A, B);
END_PROGRAM

CONFIGURATION Config0
  RESOURCE Res0 ON PLC
    TASK task0(INTERVAL := T#20ms,PRIORITY := 0);
    PROGRAM instance0 WITH task0 : program0;
  END_RESOURCE
END_CONFIGURATION

(* ---- 423-AIN.ST ---- *)
FUNCTION _BYTE_TO_INT:INT
	VAR_INPUT
		IN :	BYTE;
	END_VAR

	_BYTE_TO_INT := USINT_TO_INT(BYTE_TO_USINT(IN));
END_FUNCTION

FUNCTION _DWORD_TO_REAL:REAL
	VAR_INPUT
		IN :	DWORD;
	END_VAR

	_DWORD_TO_REAL := UDINT_TO_REAL(DWORD_TO_UDINT(IN));
END_FUNCTION

FUNCTION BIT_OF_DWORD:BOOL
	VAR_INPUT
		IN :	DWORD;
		N :	INT;
	END_VAR
	BIT_OF_DWORD := (SHR(in,n) AND DWORD#1) > DWORD#0;
END_FUNCTION

FUNCTION AIN:REAL
	VAR_INPUT
		IN :	DWORD;
		BITS :	BYTE;
		SIGN :	BYTE;
		LOW :	REAL;
		HIGH :	REAL;
	END_VAR

	VAR
		temp1 :	DWORD;
		temp2 :	DWORD;
		sx :	BOOL;
	END_VAR

	IF sign < BYTE#32 THEN
		temp1 := SHR(in, _BYTE_TO_INT(sign));
		sx := BIT_OF_DWORD(temp1,0); (* temp1.X0 *)
	ELSE
		sx := FALSE;
	END_IF;
	temp1 := SHR(DWORD#16#FFFFFFFF,32 - _BYTE_TO_INT(bits));
	temp2 := in AND temp1;
	AIN := (high - low)* _DWORD_TO_REAL(temp2) / _DWORD_TO_REAL(temp1) + low;
	IF sx THEN AIN := -AIN; END_IF;
END_FUNCTION

PROGRAM program0
  VAR
    LocalVar0 : DWORD;
	LocalVar1 : BYTE;
	LocalVar2 : BYTE;
	LocalVar3 : REAL;
	LocalVar4 : REAL;
    LocalOUT  : REAL;
  END_VAR

  LocalOUT := AIN(LocalVar0, LocalVar1, LocalVar2, LocalVar3, LocalVar4);
END_PROGRAM

CONFIGURATION Config0
  RESOURCE Res0 ON PLC
    TASK task0(INTERVAL := T#20ms,PRIORITY := 0);
    PROGRAM instance0 WITH task0 : program0;
  END_RESOURCE
END_CONFIGURATION

(* ---- 43-TANC.ST ---- *)
FUNCTION TANC:REAL

	VAR_INPUT
		X :	REAL;
	END_VAR

	IF X = 0.0 THEN
		TANC := 1.0;
	ELSE
		TANC := TAN(x) / x;
	END_IF;

END_FUNCTION

PROGRAM program0

	VAR
		X :	REAL;
		CEIL5_OUT : REAL;
	END_VAR

	CEIL5_OUT := TANC(X);

END_PROGRAM

CONFIGURATION Config0

	RESOURCE Res0 ON PLC
		TASK task0(INTERVAL := T#20ms,PRIORITY := 0);
		PROGRAM instance0 WITH task0 : program0;
	END_RESOURCE

END_CONFIGURATION

(* ---- 436-AOUT1.ST ---- *)
FUNCTION SIGN_R : BOOL
  VAR_INPUT
    IN : REAL;
  END_VAR

  SIGN_R := in < 0.0;
END_FUNCTION

FUNCTION _REAL_TO_DWORD: DWORD

  VAR_INPUT
    X :	REAL;
  END_VAR

  IF REAL_TO_DWORD(0.5) = DWORD#1 THEN
    _REAL_TO_DWORD := REAL_TO_DWORD(x);
  ELSIF X > 0.0 THEN
    _REAL_TO_DWORD := REAL_TO_DWORD(x+0.5);
  ELSIF X < 0.0 THEN
    _REAL_TO_DWORD := REAL_TO_DWORD(x-0.5);
  ELSE
    _REAL_TO_DWORD := DWORD#0;
  END_IF;
END_FUNCTION

FUNCTION AOUT1:DWORD

	VAR_INPUT
		IN :	REAL;
		BIT_0 :	INT;
		BIT_N :	INT;
		SIGN :	INT;
		LOW :	REAL;
		HIGH :	REAL;
	END_VAR

	VAR
		in2 :	REAL;
		sx :	BOOL;
	END_VAR

	IF sign < 32 THEN
		sx := sign_R(in);
		in2 := ABS(in);
	ELSE
		sx := FALSE;
		in2 := in;
	END_IF;

	in2 := LIMIT_REAL(low, in2, high);

	AOUT1 :=  SHL(_REAL_TO_DWORD((in2 - low) / (high - low) * UDINT_TO_REAL(DWORD_TO_UDINT(SHL(DWORD#2#1,bit_n - Bit_0 + 1)) - UDINT#1)),Bit_0);

	IF sx THEN AOUT1 := SHL(DWORD#2#1,sign) OR AOUT1; END_IF;

END_FUNCTION

PROGRAM program0
  VAR
    LocalVar0 : REAL;
	LocalVar1 : INT;
	LocalVar21 : INT;
	LocalVar2 : INT;
	LocalVar3 : REAL;
	LocalVar4 : REAL;
	LocalOUT  : DWORD;
  END_VAR
  	LocalOUT := AOUT1(LocalVar0, LocalVar1,LocalVar21, LocalVar2, LocalVar3,LocalVar4);
END_PROGRAM

CONFIGURATION Config0
  RESOURCE Res0 ON PLC
    TASK task0(INTERVAL := T#20ms,PRIORITY := 0);
    PROGRAM instance0 WITH task0 : program0;
  END_RESOURCE
END_CONFIGURATION

(* ---- 44-SETUP_EXTENDED_ASCII.ST ---- *)
FUNCTION SETUP_EXTENDED_ASCII:BOOL

	VAR_INPUT
		X :	BOOL;
	END_VAR

	SETUP_EXTENDED_ASCII := X OR TRUE;
END_FUNCTION

PROGRAM program0
  VAR
	X :	BOOL;
    CEIL5_OUT : BOOL;
  END_VAR

  CEIL5_OUT := SETUP_EXTENDED_ASCII(X);
END_PROGRAM

CONFIGURATION Config0

  RESOURCE Res0 ON PLC
    TASK task0(INTERVAL := T#20ms,PRIORITY := 0);
    PROGRAM instance0 WITH task0 : program0;
  END_RESOURCE
END_CONFIGURATION

(* ---- 443-SET_DT.ST ---- *)
FUNCTION _INT_TO_UDINT:UDINT
	VAR_INPUT
		IN :	INT;
	END_VAR

	_INT_TO_UDINT := DINT_TO_UDINT(INT_TO_DINT(IN));
END_FUNCTION

FUNCTION SET_DATE:UDINT

	VAR_INPUT
		YEAR :	INT;
		MONTH :	INT;
		DAY :	INT;
	END_VAR

	VAR
		count :	INT;
	END_VAR

	IF month > 2 THEN
		count := (month - 1) * 30;
		IF month > 7 THEN
			count := count + DWORD_TO_INT(SHR(DINT_TO_DWORD(INT_TO_DINT(month) - INT_TO_DINT(3)),1));
		ELSE
			count := count + DWORD_TO_INT(SHR(DINT_TO_DWORD(INT_TO_DINT(month) - INT_TO_DINT(4)),1));
		END_IF;
		IF SHL(INT_TO_WORD(year),14) = WORD#0 THEN
			count := count + 1;
		END_IF;
	ELSE
		count := (month - 1) * 31;
	END_IF;
	SET_DATE := (_INT_TO_UDINT(count + day - 1) + DWORD_TO_UDINT(SHR(UDINT_TO_DWORD(_INT_TO_UDINT(year) * UDINT#1461 - UDINT#2878169), 2))) * UDINT#86400;

END_FUNCTION

FUNCTION SET_DT:UDINT
	VAR_INPUT
		YEAR :	INT;
		MONTH :	INT;
		DAY :	INT;
		HOUR :	INT;
		MINUTE :	INT;
		SECOND :	INT;
	END_VAR

	SET_DT := SET_DATE(YEAR, MONTH, DAY) + _INT_TO_UDINT(SECOND) + _INT_TO_UDINT(MINUTE) * UDINT#60 + _INT_TO_UDINT(HOUR) * UDINT#3600;
END_FUNCTION

PROGRAM program0

	VAR
		YEAR :	INT;
		MONTH :	INT;
		DAY :	INT;
		HOUR :	INT;
		MINUTE :	INT;
		SECOND :	INT;
		CEIL5_OUT : UDINT;
	END_VAR

	CEIL5_OUT := SET_DT(YEAR, MONTH, DAY, HOUR, MINUTE, SECOND);

END_PROGRAM

CONFIGURATION Config0

	RESOURCE Res0 ON PLC
		TASK task0(INTERVAL := T#20ms,PRIORITY := 0);
		PROGRAM instance0 WITH task0 : program0;
	END_RESOURCE

END_CONFIGURATION

(* ---- 447-TRIANGLE_A.ST ---- *)
FUNCTION _REAL_TO_DINT:DINT
  VAR_INPUT
    X :	REAL;
  END_VAR

  IF REAL_TO_DINT(0.5) = DINT#1 THEN
    _REAL_TO_DINT := REAL_TO_DINT(x);
    RETURN;
  END_IF;

  IF X > 0.0 THEN
    _REAL_TO_DINT := REAL_TO_DINT(x+0.5);
  ELSIF X < 0.0 THEN
    _REAL_TO_DINT := REAL_TO_DINT(x-0.5);
  ELSE
    _REAL_TO_DINT := DINT#0;
  END_IF;
END_FUNCTION

FUNCTION FLOOR2:DINT

	VAR_INPUT
		X :	REAL;
	END_VAR

	FLOOR2 := _REAL_TO_DINT(X);
	IF DINT_TO_REAL(FLOOR2) > X THEN
		FLOOR2 := FLOOR2 - DINT#1;
	END_IF;

END_FUNCTION

FUNCTION MODR:REAL

	VAR_INPUT
		IN :	REAL;
		DIVI :	REAL;
	END_VAR

	IF divi = 0.0 THEN
		MODR := 0.0;
	ELSE
		MODR := in - DINT_TO_REAL(FLOOR2(in / divi)) * divi;
	END_IF;

END_FUNCTION

FUNCTION RAD:REAL

	VAR_INPUT
		DEG :	REAL;
	END_VAR

	Rad := modR(0.0174532925199433 * deg , 6.283185307179586476);

END_FUNCTION

FUNCTION TRIANGLE_A:REAL

	VAR_INPUT
		S1 :	REAL;
		A :	REAL;
		S2 :	REAL;
		S3 :	REAL;
	END_VAR

	IF A = 0.0 THEN
		TRIANGLE_A := SQRT((s1+s2+S3) * (s1+s2-S3) * (S2+S3-S1) * (S3+S1-S2)) * 0.25;
	ELSE
		TRIANGLE_A := S1 * S2 * SIN(RAD(A)) * 0.5;
	END_IF;

END_FUNCTION

PROGRAM program0
  VAR
	S1 :	REAL;
	A :	REAL;
	S2 :	REAL;
	S3 :	REAL;
    CEIL5_OUT : REAL;
  END_VAR

  CEIL5_OUT := TRIANGLE_A(S1, A, S2, S3);
END_PROGRAM

CONFIGURATION Config0

  RESOURCE Res0 ON PLC
    TASK task0(INTERVAL := T#20ms,PRIORITY := 0);
    PROGRAM instance0 WITH task0 : program0;
  END_RESOURCE
END_CONFIGURATION

(* ---- 45-DWORD_TO_TOD.ST ---- *)
FUNCTION DWORD_TO_TOD2:UDINT
	VAR_INPUT
		IN :	DWORD;
	END_VAR
	DWORD_TO_TOD2 := DWORD_TO_UDINT(IN);
END_FUNCTION

PROGRAM program0
  VAR
    LocalVar0 : DWORD;
	  LocalOUT  : UDINT;
  END_VAR
  	LocalOUT := DWORD_TO_TOD2(LocalVar0);
END_PROGRAM

CONFIGURATION Config0
  RESOURCE Res0 ON PLC
    TASK task0(INTERVAL := T#20ms,PRIORITY := 0);
    PROGRAM instance0 WITH task0 : program0;
  END_RESOURCE
END_CONFIGURATION

(* ---- 450-PERIOD.ST ---- *)
FUNCTION LEAP_OF_DATE:BOOL

	VAR_INPUT
		IDATE :	UDINT;
	END_VAR

	LEAP_OF_DATE := SHL(UDINT_TO_DWORD((idate + UDINT#43200) / UDINT#31557600), 30) = DWORD#16#80000000;
END_FUNCTION

FUNCTION DAY_OF_YEAR:INT
	VAR_INPUT
		IDATE :	UDINT;
	END_VAR

	DAY_OF_YEAR := UDINT_TO_INT(((idate) / UDINT#86400) MOD UDINT#1461);
	IF DAY_OF_YEAR > 729 THEN
		IF DAY_OF_YEAR > 1095 THEN DAY_OF_YEAR := DAY_OF_YEAR - 1095; ELSE DAY_OF_YEAR := DAY_OF_YEAR - 729; END_IF;
	ELSIF DAY_OF_YEAR > 364 THEN
		DAY_OF_YEAR := DAY_OF_YEAR - 364;
	ELSE
		DAY_OF_YEAR := DAY_OF_YEAR + 1;
	END_IF;
END_FUNCTION

FUNCTION PERIOD:BOOL

	VAR
		day1 :	INT;
		day2 :	INT;
		dayx :	INT;
	END_VAR

	VAR_INPUT
		D1 :	UDINT;
		Dx :	UDINT;
		D2 :	UDINT;
	END_VAR

	day1 := day_of_year(d1);
	day2 := day_of_year(d2);
	dayx := day_of_year(dx);
	IF NOT leap_of_Date(dx) AND dayx > 58 THEN dayx := dayx + 1; END_IF;
	IF NOT leap_of_Date(d1) AND day1 > 58 THEN day1 := day1 + 1; END_IF;
	IF NOT leap_of_Date(d2) AND day2 > 58 THEN day2 := day2 + 1; END_IF;

	IF day2 < day1 THEN
		(* the period spans over the new year *)
		period := dayx <= day2 OR dayx >= day1;
	ELSE
		period := dayx >= day1 AND dayx <= day2;
	END_IF;

END_FUNCTION

PROGRAM program0
	VAR
		D1 :	UDINT;
		Dx :	UDINT;
		D2 :	UDINT;

		OUT : BOOL;
	END_VAR

	OUT := PERIOD(D1, Dx, D2);
END_PROGRAM

CONFIGURATION Config0

	RESOURCE Res0 ON PLC
		TASK task0(INTERVAL := T#20ms,PRIORITY := 0);
		PROGRAM instance0 WITH task0 : program0;
	END_RESOURCE

END_CONFIGURATION

(* ---- 451-SUN_MIDDAY.ST ---- *)
FUNCTION _REAL_TO_UDINT:UDINT
	VAR_INPUT
		X :	REAL;
	END_VAR

	IF REAL_TO_UDINT(0.5) = UDINT#1 THEN
		_REAL_TO_UDINT := REAL_TO_UDINT(x);
	ELSIF X > 0.0 THEN
		_REAL_TO_UDINT := REAL_TO_UDINT(x+0.5);
	ELSIF X < 0.0 THEN
		_REAL_TO_UDINT := REAL_TO_UDINT(x-0.5);
	ELSE
		_REAL_TO_UDINT := UDINT#0;
	END_IF;

END_FUNCTION

FUNCTION HOUR_TO_TOD:UDINT

	VAR_INPUT
		IN :	REAL;
	END_VAR

	hour_to_tod := _REAL_TO_UDINT(IN * 3600000.00);

END_FUNCTION

FUNCTION DAY_OF_YEAR:INT
	VAR_INPUT
		IDATE :	DATE;
	END_VAR

	DAY_OF_YEAR := UDINT_TO_INT((DATE_TO_UDINT(idate) / UDINT#86400) MOD UDINT#1461);
	IF DAY_OF_YEAR > 729 THEN
		IF DAY_OF_YEAR > 1095 THEN DAY_OF_YEAR := DAY_OF_YEAR - 1095; ELSE DAY_OF_YEAR := DAY_OF_YEAR - 729; END_IF;
	ELSIF DAY_OF_YEAR > 364 THEN
		DAY_OF_YEAR := DAY_OF_YEAR - 364;
	ELSE
		DAY_OF_YEAR := DAY_OF_YEAR + 1;
	END_IF;
END_FUNCTION

FUNCTION SUN_MIDDAY:UDINT

	VAR_INPUT
		LON :	REAL;
		UTC :	DATE;
	END_VAR

	VAR
		T :	REAL;
		OFFSET :	REAL;
	END_VAR

	T := INT_TO_REAL(DAY_OF_YEAR(utc));
	OFFSET := -0.1752 * SIN(0.033430 * T + 0.5474) - 0.1340 * SIN(0.018234 * T - 0.1939);
	SUN_MIDDAY := HOUR_TO_TOD(12.0 - OFFSET - lon * 0.0666666666666);

END_FUNCTION

PROGRAM program0

	VAR
		LON :	REAL;
		UTC :	DATE;
		CEIL5_OUT : UDINT;
	END_VAR

	CEIL5_OUT := SUN_MIDDAY(LON, UTC);

END_PROGRAM

CONFIGURATION Config0

	RESOURCE Res0 ON PLC
		TASK task0(INTERVAL := T#20ms,PRIORITY := 0);
		PROGRAM instance0 WITH task0 : program0;
	END_RESOURCE

END_CONFIGURATION

(* ---- 454-EASTER.ST ---- *)
FUNCTION _INT_TO_UDINT:UDINT
	VAR_INPUT
		IN :	INT;
	END_VAR

	_INT_TO_UDINT := DINT_TO_UDINT(INT_TO_DINT(IN));
END_FUNCTION

FUNCTION SET_DATE:UDINT

	VAR_INPUT
		YEAR :	INT;
		MONTH :	INT;
		DAY :	INT;
	END_VAR

	VAR
		count :	INT;
	END_VAR

	IF month > 2 THEN
		count := (month - 1) * 30;
		IF month > 7 THEN
			count := count + DWORD_TO_INT(SHR(DINT_TO_DWORD(INT_TO_DINT(month) - INT_TO_DINT(3)),1));
		ELSE
			count := count + DWORD_TO_INT(SHR(DINT_TO_DWORD(INT_TO_DINT(month) - INT_TO_DINT(4)),1));
		END_IF;
		IF SHL(INT_TO_WORD(year),14) = WORD#0 THEN
			count := count + 1;
		END_IF;
	ELSE
		count := (month - 1) * 31;
	END_IF;
	SET_DATE := (_INT_TO_UDINT(count + day - 1) + DWORD_TO_UDINT(SHR(UDINT_TO_DWORD(_INT_TO_UDINT(year) * UDINT#1461 - UDINT#2878169), 2))) * UDINT#86400;

END_FUNCTION

FUNCTION EASTER:UDINT
	VAR_INPUT
		YEAR :	INT;
	END_VAR

	VAR
		b :	INT;
		c :	INT;
		oday :	INT;
	END_VAR

	b := (204 - 11 * (year MOD 19)) MOD 30;
	IF b > 27 THEN b := b - 1; END_IF;
	c := (year + WORD_TO_INT(SHR(INT_TO_WORD(year),2)) + b - 13) MOD 7;
	oday := 28 + b - c;
	IF oday > 33 THEN
		easter := set_Date(year, 4, oday - 31);
	ELSE
		easter := set_Date(year, 3, oday);
	END_IF;
END_FUNCTION

PROGRAM program0
  VAR
    LocalVar0 : INT;
	LocalOUT  : UDINT;
  END_VAR
  	LocalOUT := EASTER(LocalVar0);
END_PROGRAM

CONFIGURATION Config0
  RESOURCE Res0 ON PLC
    TASK task0(INTERVAL := T#20ms,PRIORITY := 0);
    PROGRAM instance0 WITH task0 : program0;
  END_RESOURCE
END_CONFIGURATION

(* ---- 455-DAYS_IN_MONTH.ST ---- *)
FUNCTION DAY_OF_YEAR:INT
	VAR_INPUT
		IDATE :	UDINT;
	END_VAR

	DAY_OF_YEAR := UDINT_TO_INT(((idate) / UDINT#86400) MOD UDINT#1461);
	IF DAY_OF_YEAR > 729 THEN
		IF DAY_OF_YEAR > 1095 THEN DAY_OF_YEAR := DAY_OF_YEAR - 1095; ELSE DAY_OF_YEAR := DAY_OF_YEAR - 729; END_IF;
	ELSIF DAY_OF_YEAR > 364 THEN
		DAY_OF_YEAR := DAY_OF_YEAR - 364;
	ELSE
		DAY_OF_YEAR := DAY_OF_YEAR + 1;
	END_IF;
END_FUNCTION

FUNCTION LEAP_OF_DATE:BOOL

	VAR_INPUT
		IDATE :	UDINT;
	END_VAR

	LEAP_OF_DATE := SHL(UDINT_TO_DWORD((idate + UDINT#43200) / UDINT#31557600), 30) = DWORD#16#80000000;
END_FUNCTION

FUNCTION DAYS_IN_MONTH:INT

	VAR_INPUT
		IDATE :	UDINT;
	END_VAR

	DAYS_IN_MONTH := DAY_OF_YEAR(IDATE);
	IF LEAP_OF_DATE(IDATE) THEN
		CASE DAYS_IN_MONTH OF
			32..60	:	DAYS_IN_MONTH := 29;
			92..121 :	DAYS_IN_MONTH := 30;
			153..182:	DAYS_IN_MONTH := 30;
			245..274:	DAYS_IN_MONTH := 30;
			306..335:	DAYS_IN_MONTH := 30;
		ELSE
			DAYS_IN_MONTH := 31;
		END_CASE;
	ELSE
		CASE DAYS_IN_MONTH OF
			32..59	:	DAYS_IN_MONTH := 28;
			91..120 :	DAYS_IN_MONTH := 30;
			152..181:	DAYS_IN_MONTH := 30;
			244..273:	DAYS_IN_MONTH := 30;
			305..334:	DAYS_IN_MONTH := 30;
		ELSE
			DAYS_IN_MONTH := 31;
		END_CASE;
	END_IF;

END_FUNCTION

PROGRAM program0
  VAR
    LocalVar0 : UDINT;
	LocalOUT  : INT;
  END_VAR
  	LocalOUT := DAYS_IN_MONTH(LocalVar0);
END_PROGRAM

CONFIGURATION Config0
  RESOURCE Res0 ON PLC
    TASK task0(INTERVAL := T#20ms,PRIORITY := 0);
    PROGRAM instance0 WITH task0 : program0;
  END_RESOURCE
END_CONFIGURATION

(* ---- 46-SINC.ST ---- *)
FUNCTION SINC:REAL

	VAR_INPUT
		X :	REAL;
	END_VAR

	IF X = 0.0 THEN
		SINC := 1.0;
	ELSE
		SINC := SIN(x) / x;
	END_IF;

END_FUNCTION

PROGRAM program0

	VAR
		X :	REAL;
		CEIL5_OUT : REAL;
	END_VAR

  	CEIL5_OUT := SINC(X);

END_PROGRAM

CONFIGURATION Config0

	RESOURCE Res0 ON PLC
		TASK task0(INTERVAL := T#20ms,PRIORITY := 0);
		PROGRAM instance0 WITH task0 : program0;
	END_RESOURCE

END_CONFIGURATION

(* ---- 468-AOUT.ST ---- *)
FUNCTION _DWORD_TO_REAL:REAL
	VAR_INPUT
		IN :	DWORD;
	END_VAR

	_DWORD_TO_REAL := UDINT_TO_REAL(DWORD_TO_UDINT(IN));
END_FUNCTION

FUNCTION SIGN_R : BOOL
  VAR_INPUT
    IN : REAL;
  END_VAR
  SIGN_R := in < 0.0;
END_FUNCTION

FUNCTION _REAL_TO_DWORD: DWORD

  VAR_INPUT
    X :	REAL;
  END_VAR

  IF REAL_TO_DWORD(0.5) = DWORD#1 THEN
    _REAL_TO_DWORD := REAL_TO_DWORD(x);
  ELSIF X > 0.0 THEN
    _REAL_TO_DWORD := REAL_TO_DWORD(x+0.5);
  ELSIF X < 0.0 THEN
    _REAL_TO_DWORD := REAL_TO_DWORD(x-0.5);
  ELSE
    _REAL_TO_DWORD := DWORD#0;
  END_IF;
END_FUNCTION

FUNCTION _BYTE_TO_INT:INT
	VAR_INPUT
		IN :	BYTE;
	END_VAR

	_BYTE_TO_INT := USINT_TO_INT(BYTE_TO_USINT(IN));
END_FUNCTION

FUNCTION AOUT:DWORD
	VAR_INPUT
		IN :	REAL;
		BITS :	BYTE;
		SIGN :	BYTE;
		LOW :	REAL;
		HIGH :	REAL;
	END_VAR

	VAR
		in2 :	REAL;
		sx :	BOOL;
	END_VAR

	IF sign < BYTE#32 THEN
		sx := sign_R(in);
		in2 := ABS(in);
	ELSE
		in2 := in;
	END_IF;

	in2 := LIMIT(low, in2, high);

	Aout := _REAL_TO_DWORD((in2 - low) / (high - low) * (_DWORD_TO_REAL(SHL(DWORD#2#1,_BYTE_TO_INT(bits))) - 1.0)   );
	IF sx THEN Aout := SHL(DWORD#2#1,_BYTE_TO_INT(sign)) OR Aout; END_IF;

END_FUNCTION

PROGRAM program0
  VAR
    LocalVar0 : REAL;
	LocalVar1 : BYTE;
	LocalVar2 : BYTE;
	LocalVar3 : REAL;
	LocalVar4 : REAL;
	LocalOUT  : DWORD;
  END_VAR
  	LocalOUT := AOUT(LocalVar0, LocalVar1, LocalVar2, LocalVar3,LocalVar4);
END_PROGRAM

CONFIGURATION Config0
  RESOURCE Res0 ON PLC
    TASK task0(INTERVAL := T#20ms,PRIORITY := 0);
    PROGRAM instance0 WITH task0 : program0;
  END_RESOURCE
END_CONFIGURATION

(* ---- 47-DATE_TO_DWORD.ST ---- *)
FUNCTION DATE_TO_DWORD2:DWORD
	VAR_INPUT
		IN :	UDINT;
	END_VAR

	DATE_TO_DWORD2 := UDINT_TO_DWORD(IN);
END_FUNCTION

PROGRAM program0
  VAR
    LocalVar0 : UDINT;
	LocalOUT  : DWORD;
  END_VAR
  	LocalOUT := DATE_TO_DWORD2(LocalVar0);
END_PROGRAM

CONFIGURATION Config0
  RESOURCE Res0 ON PLC
    TASK task0(INTERVAL := T#20ms,PRIORITY := 0);
    PROGRAM instance0 WITH task0 : program0;
  END_RESOURCE
END_CONFIGURATION

(* ---- 470-SCALE_X8.ST ---- *)
FUNCTION SCALE_X8:REAL

	VAR_INPUT
		IN1 :	BOOL;
		IN2 :	BOOL;
		IN3 :	BOOL;
		IN4 :	BOOL;
		IN5 :	BOOL;
		IN6 :	BOOL;
		IN7 :	BOOL;
		IN8 :	BOOL;
		K :	REAL;
		O :	REAL;
		IN1_MIN :	REAL;
		IN1_MAX :	REAL;
		IN2_MIN :	REAL;
		IN2_MAX :	REAL;
		IN3_MIN :	REAL;
		IN3_MAX :	REAL;
		IN4_MIN :	REAL;
		IN4_MAX :	REAL;
		IN5_MIN :	REAL;
		IN5_MAX :	REAL;
		IN6_MIN :	REAL;
		IN6_MAX :	REAL;
		IN7_MIN :	REAL;
		IN7_MAX :	REAL;
		IN8_MIN :	REAL;
		IN8_MAX :	REAL;
	END_VAR

	SCALE_X8 := (SEL(IN1,IN1_MIN, IN1_MAX)+ SEL(IN2,IN2_MIN, IN2_MAX)+SEL(IN3,IN3_MIN, IN3_MAX)+ SEL(IN4,IN4_MIN, IN4_MAX)
					+SEL(IN5,IN5_MIN, IN5_MAX)+ SEL(IN6,IN6_MIN, IN6_MAX)+SEL(IN7,IN7_MIN, IN7_MAX)+ SEL(IN8,IN8_MIN, IN8_MAX))*k + o;

END_FUNCTION

PROGRAM program0

  	VAR
		IN1 :	BOOL;
		IN2 :	BOOL;
		IN3 :	BOOL;
		IN4 :	BOOL;
		IN5 :	BOOL;
		IN6 :	BOOL;
		IN7 :	BOOL;
		IN8 :	BOOL;
		K :	REAL;
		O :	REAL;
		IN1_MIN :	REAL;
		IN1_MAX :	REAL;
		IN2_MIN :	REAL;
		IN2_MAX :	REAL;
		IN3_MIN :	REAL;
		IN3_MAX :	REAL;
		IN4_MIN :	REAL;
		IN4_MAX :	REAL;
		IN5_MIN :	REAL;
		IN5_MAX :	REAL;
		IN6_MIN :	REAL;
		IN6_MAX :	REAL;
		IN7_MIN :	REAL;
		IN7_MAX :	REAL;
		IN8_MIN :	REAL;
		IN8_MAX :	REAL;
		CEIL5_OUT : REAL;
  	END_VAR

  	CEIL5_OUT := SCALE_X8(IN1, IN2, IN3, IN4, IN5, IN6, IN7, IN8, K, O, IN1_MIN, IN1_MAX, IN2_MIN, IN2_MAX, IN3_MIN, IN3_MAX, IN4_MIN, IN4_MAX, IN5_MIN, IN5_MAX, IN6_MIN, IN6_MAX, IN7_MIN, IN7_MAX, IN8_MIN, IN8_MAX);
END_PROGRAM

CONFIGURATION Config0

	RESOURCE Res0 ON PLC
		TASK task0(INTERVAL := T#20ms,PRIORITY := 0);
		PROGRAM instance0 WITH task0 : program0;
	END_RESOURCE

END_CONFIGURATION

(* ---- 48-TIME_TO_TOD.ST ---- *)
FUNCTION TIME_TO_TOD:UDINT

	VAR_INPUT
		IN :	TIME;
	END_VAR

	TIME_TO_TOD := DWORD_TO_UDINT(TIME_TO_DWORD(IN));
END_FUNCTION

PROGRAM program0
  VAR
	IN :	TIME;
    CEIL5_OUT : UDINT;
  END_VAR

  CEIL5_OUT := TIME_TO_TOD(IN);
END_PROGRAM

CONFIGURATION Config0

  RESOURCE Res0 ON PLC
    TASK task0(INTERVAL := T#20ms,PRIORITY := 0);
    PROGRAM instance0 WITH task0 : program0;
  END_RESOURCE
END_CONFIGURATION

(* ---- 481-RND.ST ---- *)
FUNCTION CEIL:INT

	VAR_INPUT
		X :	REAL;
	END_VAR

	CEIL := REAL_TO_INT(x);
	IF INT_TO_REAL(CEIL) < X THEN
			CEIL := CEIL + 1;
	END_IF;

END_FUNCTION

FUNCTION BIT_OF_DWORD : BOOL

	VAR_INPUT
		IN : DWORD;
		N : INT;
	END_VAR

	BIT_OF_DWORD := (SHR(in,N) AND 16#00000001) > 0;

END_FUNCTION

FUNCTION EXPN:REAL

	VAR_INPUT
		X :	REAL;
		N :	INT;
	END_VAR

	VAR
		N_word :	WORD;
		X_tmp :	REAL;
		sign :	BOOL;
	END_VAR

	N_word := INT_TO_WORD(N);
	X_tmp := X;
	sign := BIT_OF_DWORD(WORD_TO_DWORD(N_word),15);
	N_word := INT_TO_WORD(ABS(N));
	IF BIT_OF_DWORD(WORD_TO_DWORD(N_word),0) THEN expn := X_tmp; ELSE expn := 1.0; END_IF;    (* N_word.X0 *)
	N_word := SHR(N_word,1);
	WHILE N_word > WORD#0 DO
		X_tmp := X_tmp * X_tmp;
		IF BIT_OF_DWORD(WORD_TO_DWORD(N_word),0) THEN expn := expn * X_tmp; END_IF;       (* N_word.X0 *)
		N_word := SHR(N_word,1);
	END_WHILE;
	IF sign THEN EXPN := 1.0 / EXPN; END_IF;

END_FUNCTION

FUNCTION _REAL_TO_DINT:DINT
	VAR_INPUT
		X :	REAL;
	END_VAR

	IF REAL_TO_DINT(0.5) = DINT#1 THEN
		_REAL_TO_DINT := REAL_TO_DINT(x);
		RETURN;
	END_IF;

	IF X > 0.0 THEN
		_REAL_TO_DINT := REAL_TO_DINT(x+0.5);
	ELSIF X < 0.0 THEN
		_REAL_TO_DINT := REAL_TO_DINT(x-0.5);
	ELSE
		_REAL_TO_DINT := DINT#0;
	END_IF;
END_FUNCTION

FUNCTION RND:REAL

	VAR_INPUT
		X :	REAL;
		N :	INT;
	END_VAR

	VAR
		M :	REAL;
	END_VAR

	IF X = 0.0 THEN
		RND := 0.0;
	ELSE
		M := EXPN(10.0,N - CEIL(LOG(ABS(X))));
		RND := DINT_TO_REAL(_REAL_TO_DINT(X * M)) / M;
	END_IF;

END_FUNCTION

PROGRAM program0
	VAR
		IN : REAL;
		N :	INT;
		X :	REAL;
	END_VAR
		X := RND(IN, N);
END_PROGRAM

CONFIGURATION Config0

	RESOURCE Res0 ON PLC
		TASK task0(INTERVAL := T#20ms,PRIORITY := 0);
		PROGRAM instance0 WITH task0 : program0;
	END_RESOURCE

END_CONFIGURATION

(* ---- 485-INI_PARSER_FILE_DEMO.ST ---- *)
PROGRAM INI_PARSER_FILE_DEMO

	VAR

	END_VAR

	VAR_EXTERNAL

	END_VAR

	VAR
		SMTP_SERVER :	STRING;
		SMTP_FROM :	STRING;
		STATION_NAME :	STRING;
		STATION_IP :	STRING;
	END_VAR

	VAR
		IPF :	INI_PARSER_FILE;
		FS :	FILE_SERVER;
		FSD :	oscat_FILE_SERVER_DATA;
		PT :	oscat_NETWORK_BUFFER;
		section :	INT;
		filename :	STRING;
		key :	oscat_STRING250;
		value :	oscat_STRING250;
		str :	oscat_STRING250;
		step :	INT;
		result :	BYTE;
		offset :	UDINT;
		run :	BYTE;
		done :	BOOL;
	END_VAR

	CASE step OF

	00:	IF NOT done THEN
			filename := 'config.ini';
			offset := UDINT#0;
			str := '';
			run := BYTE#3;
			step := 50;
		END_IF;

	50:	IF run = BYTE#0 THEN

			run := BYTE#3;

			IF result = BYTE#1 THEN
				IF EQ_STRING(key,'Station') THEN
					section := 1;
				ELSIF EQ_STRING(key,'SMTP') THEN
					section := 2;

				ELSE
					section := 0;
				END_IF;

			ELSIF result = BYTE#2 AND section > 0 THEN

				CASE section OF

				1:
					IF EQ_STRING(key,'NAME') THEN
						STATION_NAME := value;
					ELSIF EQ_STRING(key,'IP') THEN
						STATION_IP := value;
					END_IF;

				2:
					IF EQ_STRING(key,'SERVER') THEN
						SMTP_SERVER := value;
					ELSIF EQ_STRING(key,'FROM') THEN
						SMTP_FROM := value;
					END_IF;

				END_CASE;

			ELSIF result = BYTE#10 THEN
				run := BYTE#0;
				FSD.MODE := BYTE#5;
				step := 30;
			END_IF;
		END_IF;

	30:	IF FSD.MODE = BYTE#0 THEN
			step := 0;
			done := TRUE;
		END_IF;

	END_CASE;

	IPF(FILENAME:=FILENAME,FSD:=FSD,STR:=str,RUN:=run,OFFSET:=offset,KEY:=key,VALUE:=value,PT:=PT);
	FILENAME:=IPF.FILENAME;
	FSD:=IPF.FSD;
	str:=IPF.STR;
	run:=IPF.RUN;
	offset:=IPF.OFFSET;
	key:=IPF.KEY;
	value:=IPF.VALUE;
	PT:=IPF.PT;
	result:=IPF.RESULT;

	FS(FSD:=FSD,PT:=PT);
	FSD:=FS.FSD;
	PT:=FS.PT;

END_PROGRAM

(* ---- 49-DWORD_TO_DATE.ST ---- *)
FUNCTION DWORD_TO_DATE2:UDINT
	VAR_INPUT
		IN :	DWORD;
	END_VAR
	DWORD_TO_DATE2 := DWORD_TO_UDINT(IN);
END_FUNCTION

PROGRAM program0
  VAR
    LocalVar0 : DWORD;
	LocalOUT  : UDINT;
  END_VAR
  	LocalOUT := DWORD_TO_DATE2(LocalVar0);
END_PROGRAM

CONFIGURATION Config0
  RESOURCE Res0 ON PLC
    TASK task0(INTERVAL := T#20ms,PRIORITY := 0);
    PROGRAM instance0 WITH task0 : program0;
  END_RESOURCE
END_CONFIGURATION

(* ---- 492-INI_PARSER_BUF_DEMO.ST ---- *)
PROGRAM INI_PARSER_BUF_DEMO

	VAR

	END_VAR

	VAR_EXTERNAL

	END_VAR

	VAR
		SMTP_SERVER :	STRING;
		SMTP_FROM :	STRING;
		STATION_NAME :	STRING;
		STATION_IP :	STRING;
	END_VAR

	VAR
		IPB :	INI_PARSER_BUF;
		FS :	FILE_SERVER;
		FSD :	oscat_FILE_SERVER_DATA;
		PT :	oscat_NETWORK_BUFFER;
		section :	INT;
		key :	oscat_STRING250;
		value :	oscat_STRING250;
		str :	oscat_STRING250;
		step :	INT;
		result :	BYTE;
		offset :	UDINT;
		run :	BYTE;
		done :	BOOL;
	END_VAR

	CASE step OF

	00:	IF NOT done then
			FSD.FILENAME := 'config.ini';
			FSD.MODE := BYTE#1;
			FSD.OFFSET := UDINT#0;
			FSD.AUTO_CLOSE := T#0s;
			PT.SIZE := UINT#65535;
			step := 10;
		END_IF;

	10:	IF FSD.MODE = BYTE#0 THEN
			offset := UDINT#0;
			str := '';
			run := BYTE#3;
			step := 50;
		END_IF;

	50:	IF run = BYTE#0 THEN
			run := BYTE#3;

			IF result = BYTE#1 THEN
				IF EQ_STRING(key,'Station') THEN
					section := 1;
				ELSIF EQ_STRING(key,'SMTP') THEN
					section := 2;

				ELSE
					section := 0;
				END_IF;

			ELSIF result = BYTE#2 AND section > 0 THEN

				CASE section OF

				1:
					IF EQ_STRING(key,'NAME') THEN
						STATION_NAME := value;
					ELSIF EQ_STRING(key,'IP') THEN
						STATION_IP := value;
					END_IF;

				2:
					IF EQ_STRING(key,'SERVER') THEN
						SMTP_SERVER := value;
					ELSIF EQ_STRING(key,'FROM') THEN
						SMTP_FROM := value;
					END_IF;

				END_CASE;

			ELSIF result = BYTE#10 THEN
				run := BYTE#0;
				FSD.MODE := BYTE#5;
				step := 80;
			END_IF;
		END_IF;

	80:	IF FSD.MODE = BYTE#0 THEN
			done := TRUE;
			step := 0;
		END_IF;

	END_CASE;

	IPB(STR:=str,RUN:=run,OFFSET:=offset,KEY:=key,VALUE:=value,PT:=PT);
	str:=IPB.STR;
	run:=IPB.RUN;
	offset:=IPB.OFFSET;
	key:=IPB.KEY;
	value:=IPB.VALUE;
	PT:=IPB.PT;
	result:=IPB.RESULT;

	FS(FSD:=FSD,PT:=PT);
	FSD:=FS.FSD;
	PT:=FS.PT;

END_PROGRAM

(* ---- 5-NEGX.ST ---- *)
FUNCTION NEGX:REAL

	VAR_INPUT
		X :	REAL;
	END_VAR

	NEGX := -X;

END_FUNCTION

PROGRAM program0
	VAR
		_X : REAL;
		OUT : REAL;
	END_VAR

	OUT := NEGX(_X);
END_PROGRAM

CONFIGURATION Config0

	RESOURCE Res0 ON PLC
		TASK task0(INTERVAL := T#20ms,PRIORITY := 0);
		PROGRAM instance0 WITH task0 : program0;
	END_RESOURCE

END_CONFIGURATION

(* ---- 50-MIX.ST ---- *)
FUNCTION MIX:REAL

	VAR_INPUT
		A :	REAL;
		B :	REAL;
		M :	REAL;
	END_VAR

	MIX := (1.0 - M) * A + M * B;

END_FUNCTION

PROGRAM program0
	VAR
		A :	REAL;
		B :	REAL;
		M :	REAL;

		OUT : REAL;
	END_VAR

	OUT := MIX(A, B, M);

END_PROGRAM

CONFIGURATION Config0

	RESOURCE Res0 ON PLC
		TASK task0(INTERVAL := T#20ms,PRIORITY := 0);
		PROGRAM instance0 WITH task0 : program0;
	END_RESOURCE

END_CONFIGURATION

(* ---- 501-SCALE_B8.ST ---- *)
FUNCTION _BYTE_TO_REAL:REAL
	VAR_INPUT
		IN :	BYTE;
	END_VAR

	_BYTE_TO_REAL := USINT_TO_REAL(BYTE_TO_USINT(IN));
END_FUNCTION

FUNCTION SCALE_B8:REAL
	VAR_INPUT
		IN1 :	BYTE;
		IN2 :	BYTE;
		IN3 :	BYTE;
		IN4 :	BYTE;
		IN5 :	BYTE;
		IN6 :	BYTE;
		IN7 :	BYTE;
		IN8 :	BYTE;
		K :	REAL;
		O :	REAL;
		IN1_MIN :	REAL;
		IN1_MAX :	REAL;
		IN2_MIN :	REAL;
		IN2_MAX :	REAL;
		IN3_MIN :	REAL;
		IN3_MAX :	REAL;
		IN4_MIN :	REAL;
		IN4_MAX :	REAL;
		IN5_MIN :	REAL;
		IN5_MAX :	REAL;
		IN6_MIN :	REAL;
		IN6_MAX :	REAL;
		IN7_MIN :	REAL;
		IN7_MAX :	REAL;
		IN8_MIN :	REAL;
		IN8_MAX :	REAL;
	END_VAR

	SCALE_B8 := 	(((in1_max - in1_min)* _BYTE_TO_REAL(in1) + (in2_max - in2_min)* _BYTE_TO_REAL(in2) + (in3_max - in3_min)* _BYTE_TO_REAL(in3) + (in4_max - in4_min)* _BYTE_TO_REAL(in4) +
					(in5_max - in5_min)* _BYTE_TO_REAL(in5) + (in6_max - in6_min)* _BYTE_TO_REAL(in6) + (in7_max - in7_min)* _BYTE_TO_REAL(in7) + (in8_max - in8_min)* _BYTE_TO_REAL(in8)) * 0.003921569
					+ in1_min + in2_min + in3_min + in4_min + in5_min + in6_min + in7_min + in8_min) * K + O;

END_FUNCTION

PROGRAM program0
  	VAR
		IN1 :	BYTE;
		IN2 :	BYTE;
		IN3 :	BYTE;
		IN4 :	BYTE;
		IN5 :	BYTE;
		IN6 :	BYTE;
		IN7 :	BYTE;
		IN8 :	BYTE;
		K :	REAL;
		O :	REAL;
		IN1_MIN :	REAL;
		IN1_MAX :	REAL;
		IN2_MIN :	REAL;
		IN2_MAX :	REAL;
		IN3_MIN :	REAL;
		IN3_MAX :	REAL;
		IN4_MIN :	REAL;
		IN4_MAX :	REAL;
		IN5_MIN :	REAL;
		IN5_MAX :	REAL;
		IN6_MIN :	REAL;
		IN6_MAX :	REAL;
		IN7_MIN :	REAL;
		IN7_MAX :	REAL;
		IN8_MIN :	REAL;
		IN8_MAX :	REAL;
		CEIL5_OUT : REAL;
  	END_VAR

  	CEIL5_OUT := SCALE_B8(IN1, IN2, IN3, IN4, IN5, IN6, IN7, IN8, K, O, IN1_MIN, IN1_MAX, IN2_MIN, IN2_MAX, IN3_MIN, IN3_MAX, IN4_MIN, IN4_MAX, IN5_MIN, IN5_MAX, IN6_MIN, IN6_MAX, IN7_MIN, IN7_MAX, IN8_MIN, IN8_MAX);

	END_PROGRAM

CONFIGURATION Config0

	RESOURCE Res0 ON PLC
		TASK task0(INTERVAL := T#20ms,PRIORITY := 0);
		PROGRAM instance0 WITH task0 : program0;
	END_RESOURCE

END_CONFIGURATION

(* ---- 51-_BYTE_TO_INT.ST ---- *)
FUNCTION _BYTE_TO_INT:INT
	VAR_INPUT
		IN :	BYTE;
	END_VAR

	_BYTE_TO_INT := USINT_TO_INT(BYTE_TO_USINT(IN));
END_FUNCTION

PROGRAM program0
  VAR
    LocalVar0 : BYTE;
	LocalOUT  : INT;
  END_VAR

  LocalOUT := _BYTE_TO_INT(LocalVar0);
END_PROGRAM

CONFIGURATION Config0
  RESOURCE Res0 ON PLC
    TASK task0(INTERVAL := T#20ms,PRIORITY := 0);
    PROGRAM instance0 WITH task0 : program0;
  END_RESOURCE
END_CONFIGURATION

(* ---- 511-DST.ST ---- *)
FUNCTION _INT_TO_UDINT:UDINT
	VAR_INPUT
		IN :	INT;
	END_VAR

	_INT_TO_UDINT := DINT_TO_UDINT(INT_TO_DINT(IN));
END_FUNCTION

FUNCTION YEAR_OF_DATE:INT
	VAR_INPUT
		IDATE :	UDINT;
	END_VAR

	YEAR_OF_DATE := UDINT_TO_INT((idate+UDINT#43200) / UDINT#31557600 + UDINT#1970);
END_FUNCTION

FUNCTION DT_TO_DATE2:UDINT

	VAR_INPUT
		IN :	UDINT;
	END_VAR

	DT_TO_DATE2 := (IN / UDINT#86400) * UDINT#86400;
END_FUNCTION

FUNCTION SET_DATE:UDINT

	VAR_INPUT
		YEAR :	INT;
		MONTH :	INT;
		DAY :	INT;
	END_VAR

	VAR
		count :	INT;
	END_VAR

	IF month > 2 THEN
		count := (month - 1) * 30;
		IF month > 7 THEN
			count := count + DWORD_TO_INT(SHR(DINT_TO_DWORD(INT_TO_DINT(month) - INT_TO_DINT(3)),1));
		ELSE
			count := count + DWORD_TO_INT(SHR(DINT_TO_DWORD(INT_TO_DINT(month) - INT_TO_DINT(4)),1));
		END_IF;
		IF SHL(INT_TO_WORD(year),14) = WORD#0 THEN
			count := count + 1;
		END_IF;
	ELSE
		count := (month - 1) * 31;
	END_IF;
	SET_DATE := (_INT_TO_UDINT(count + day - 1) + DWORD_TO_UDINT(SHR(UDINT_TO_DWORD(_INT_TO_UDINT(year) * UDINT#1461 - UDINT#2878169), 2))) * UDINT#86400;

END_FUNCTION

FUNCTION SET_DT:UDINT

	VAR_INPUT
		YEAR :	INT;
		MONTH :	INT;
		DAY :	INT;
		HOUR :	INT;
		MINUTE :	INT;
		SECOND :	INT;
	END_VAR

	SET_DT := SET_DATE(YEAR, MONTH, DAY) + _INT_TO_UDINT(SECOND) + _INT_TO_UDINT(MINUTE) * UDINT#60 + _INT_TO_UDINT(HOUR) * UDINT#3600;

END_FUNCTION

FUNCTION DST:BOOL
	VAR_INPUT
		UTC :	UDINT;
	END_VAR

	VAR
		yr :	INT;
		yr4 :	UDINT;
		ltc :	UDINT;
		idate :	UDINT;
	END_VAR

	yr := YEAR_OF_DATE(DT_TO_DATE2(UTC));
	ltc := UTC;
	idate := SET_DT(yr, 3, 31, 1, 0, 0);
	yr4 := DWORD_TO_UDINT(SHR(INT_TO_DWORD(5 * yr), 2)) + UDINT#1;
	DST := (idate - ((yr4 + UDINT#3) MOD UDINT#7) * UDINT#86400 <= ltc) AND (idate + (UDINT#214 - (yr4) MOD UDINT#7) * UDINT#86400 > ltc);
END_FUNCTION

PROGRAM program0
	VAR
		UTC :	UDINT;
		CEIL5_OUT : BOOL;
	END_VAR

  CEIL5_OUT := DST(UTC);

END_PROGRAM

CONFIGURATION Config0
	RESOURCE Res0 ON PLC
		TASK task0(INTERVAL := T#20ms,PRIORITY := 0);
		PROGRAM instance0 WITH task0 : program0;
	END_RESOURCE
END_CONFIGURATION

(* ---- 52-BFT_TO_MS.ST ---- *)
FUNCTION BFT_TO_MS:REAL
	VAR_INPUT
		BFT :	INT;
	END_VAR

	BFT_TO_MS := EXPT(INT_TO_REAL(BFT), 1.5) * 0.836;

END_FUNCTION

PROGRAM program0
  VAR
    LocalVar0 : INT;
    LocalOUT  : REAL;
  END_VAR

  LocalOUT := BFT_TO_MS(LocalVar0);
END_PROGRAM

CONFIGURATION Config0
  RESOURCE Res0 ON PLC
    TASK task0(INTERVAL := T#20ms,PRIORITY := 0);
    PROGRAM instance0 WITH task0 : program0;
  END_RESOURCE
END_CONFIGURATION

(* ---- 520-WORK_WEEK.ST ---- *)
FUNCTION LEAP_YEAR:BOOL

  VAR_INPUT
    YEAR :	INT;
  END_VAR

  IF (year MOD INT#400) = INT#00 THEN
    leap_year := TRUE;
  ELSIF (year MOD INT#100) = INT#00 THEN
    leap_year := FALSE;
  ELSIF (year MOD INT#04) = INT#00 THEN
    leap_year := TRUE;
  ELSE
    leap_year := FALSE;
  END_IF;

END_FUNCTION

FUNCTION DAY_OF_WEEK:INT

	VAR_INPUT
		IDATE :	UDINT;
	END_VAR

	DAY_OF_WEEK := UDINT_TO_INT((idate / UDINT#86400 + UDINT#3) MOD UDINT#7) + INT#01;

END_FUNCTION

FUNCTION YEAR_OF_DATE:INT
	VAR_INPUT
		IDATE :	UDINT;
	END_VAR

	YEAR_OF_DATE := UDINT_TO_INT((idate+UDINT#43200) / UDINT#31557600 + UDINT#1970);
END_FUNCTION

FUNCTION _INT_TO_UDINT:UDINT
	VAR_INPUT
		IN :	INT;
	END_VAR

	_INT_TO_UDINT := DINT_TO_UDINT(INT_TO_DINT(IN));
END_FUNCTION

FUNCTION YEAR_BEGIN:UDINT
	VAR_INPUT
		Y :	INT;
	END_VAR
	year_begin := DWORD_TO_UDINT(SHR(UDINT_TO_DWORD(_INT_TO_UDINT(y) * UDINT#1461 - UDINT#2878169),2))*UDINT#86400;

END_FUNCTION

FUNCTION WORK_WEEK:INT

	VAR_INPUT
		IDATE :	UDINT;
	END_VAR

	VAR
		d1 :	UDINT;
		w1 :	INT;
		ds :	UDINT;
		yr :	INT;
		w31 :	INT;
		w01 :	INT;
		wm :	INT;
	END_VAR

	yr := YEAR_OF_DATE(idate);
	d1 := year_begin(yr);
	w1 := DAY_OF_WEEK(d1);
	IF w1 < 5 THEN
		ds := d1 - _INT_TO_UDINT(w1+6) * UDINT#86400;
	ELSE
		ds := d1 + _INT_TO_UDINT(1-w1) * UDINT#86400;
	END_IF;

	work_week := UDINT_TO_INT((idate - ds) / UDINT#604800);

	IF work_week = 0 THEN
		IF w1 > 1 THEN w31 := w1 - 1; ELSE W31 := 7; END_IF;
		IF leap_year(yr - 1) THEN IF w31 > 1 THEN w01 := W31 - 1; ELSE w1 := 7; END_IF; END_IF;
		WORK_WEEK := 52 + BOOL_TO_INT(w31 = 4 OR w01 = 4);
	ELSE
		IF leap_year(yr) THEN
			IF w1 < 7 THEN w31 := w1 + 1; ELSE w31 := 1; END_IF;
		ELSE
			w31 := w1;
		END_IF;
		wm := 52 + BOOL_TO_INT(w31 = 4 OR w1 = 4);
		IF work_week > wm THEN work_week := 1; END_IF;
	END_IF;

END_FUNCTION

PROGRAM program0
  VAR
    Y : UDINT;
    CEIL5_OUT : INT;
  END_VAR

  CEIL5_OUT := WORK_WEEK(Y);
END_PROGRAM

CONFIGURATION Config0

  RESOURCE Res0 ON PLC
    TASK task0(INTERVAL := T#20ms,PRIORITY := 0);
    PROGRAM instance0 WITH task0 : program0;
  END_RESOURCE
END_CONFIGURATION

(* ---- 528-DAY_OF_MONTH.ST ---- *)
FUNCTION LEAP_OF_DATE:BOOL

	VAR_INPUT
		IDATE :	UDINT;
	END_VAR

	LEAP_OF_DATE := SHL(UDINT_TO_DWORD((idate + UDINT#43200) / UDINT#31557600), 30) = DWORD#16#80000000;

END_FUNCTION

FUNCTION DAY_OF_YEAR:INT
	VAR_INPUT
		IDATE :	DATE;
	END_VAR

	DAY_OF_YEAR := UDINT_TO_INT((DATE_TO_UDINT(idate) / UDINT#86400) MOD UDINT#1461);
	IF DAY_OF_YEAR > 729 THEN
		IF DAY_OF_YEAR > 1095 THEN DAY_OF_YEAR := DAY_OF_YEAR - 1095; ELSE DAY_OF_YEAR := DAY_OF_YEAR - 729; END_IF;
	ELSIF DAY_OF_YEAR > 364 THEN
		DAY_OF_YEAR := DAY_OF_YEAR - 364;
	ELSE
		DAY_OF_YEAR := DAY_OF_YEAR + 1;
	END_IF;
END_FUNCTION

FUNCTION DAY_OF_MONTH:INT
	VAR_INPUT
		IDATE :	DATE;
	END_VAR

	day_of_month := day_of_year(idate);

	IF leap_of_Date(DATE_TO_UDINT(idate)) THEN
		CASE day_of_month OF
			32..60	:	day_of_month := day_of_month - 31;
			61..91	:	day_of_month := day_of_month - 60;
			92..121 :	day_of_month := day_of_month - 91;
			122..152:	day_of_month := day_of_month - 121;
			153..182:	day_of_month := day_of_month - 152;
			183..213:	day_of_month := day_of_month - 182;
			214..244:	day_of_month := day_of_month - 213;
			245..274:	day_of_month := day_of_month - 244;
			275..305:	day_of_month := day_of_month - 274;
			306..335:	day_of_month := day_of_month - 305;
			336..366:	day_of_month := day_of_month - 335;
		END_CASE;
	ELSE
		CASE day_of_month OF
			32..59	:	day_of_month := day_of_month - 31;
			60..90	:	day_of_month := day_of_month - 59;
			91..120 :	day_of_month := day_of_month - 90;
			121..151:	day_of_month := day_of_month - 120;
			152..181:	day_of_month := day_of_month - 151;
			182..212:	day_of_month := day_of_month - 181;
			213..243:	day_of_month := day_of_month - 212;
			244..273:	day_of_month := day_of_month - 243;
			274..304:	day_of_month := day_of_month - 273;
			305..334:	day_of_month := day_of_month - 304;
			335..365:	day_of_month := day_of_month - 334;
		END_CASE;
	END_IF;

END_FUNCTION

PROGRAM program0
  VAR
    LocalVar0 : DATE;
	LocalOUT  : INT;
  END_VAR
  	LocalOUT := DAY_OF_MONTH(LocalVar0);
END_PROGRAM

CONFIGURATION Config0
  RESOURCE Res0 ON PLC
    TASK task0(INTERVAL := T#20ms,PRIORITY := 0);
    PROGRAM instance0 WITH task0 : program0;
  END_RESOURCE
END_CONFIGURATION

(* ---- 53-SECOND.ST ---- *)
FUNCTION SECOND:REAL

	VAR_INPUT
		ITOD :	UDINT;
	END_VAR

	second := UDINT_TO_REAL(itod MOD UDINT#60000) / REAL#1000.00;

END_FUNCTION

PROGRAM program0
  VAR
    ITOD :	UDINT;
    CEIL5_OUT : REAL;
  END_VAR

  CEIL5_OUT := SECOND(ITOD);
END_PROGRAM

CONFIGURATION Config0

	RESOURCE Res0 ON PLC
		TASK task0(INTERVAL := T#20ms,PRIORITY := 0);
		PROGRAM instance0 WITH task0 : program0;
	END_RESOURCE

END_CONFIGURATION

(* ---- 54-TIME_TO_REAL.ST ---- *)
FUNCTION TIME_TO_REAL1:REAL

VAR_INPUT
	X :	TIME;
END_VAR

TIME_TO_REAL1 := UDINT_TO_REAL(DINT_TO_UDINT(TIME_TO_DINT(X)));
END_FUNCTION

PROGRAM program0
  VAR
	X :	TIME;
    CEIL5_OUT : REAL;
  END_VAR

  CEIL5_OUT := TIME_TO_REAL1(X);
END_PROGRAM

CONFIGURATION Config0

  RESOURCE Res0 ON PLC
    TASK task0(INTERVAL := T#20ms,PRIORITY := 0);
    PROGRAM instance0 WITH task0 : program0;
  END_RESOURCE
END_CONFIGURATION

(* ---- 55-INT_TO_BCDC.ST ---- *)
FUNCTION INT_TO_BCDC:BYTE

	VAR_INPUT
		IN :	INT;
	END_VAR

	INT_TO_BCDC := SHL(INT_TO_BYTE(IN / INT#10),4) OR INT_TO_BYTE(in MOD INT#10);

END_FUNCTION

PROGRAM program0

	VAR
		IN :	INT;
		OUT : BYTE;
	END_VAR

	OUT := INT_TO_BCDC(IN);

END_PROGRAM

CONFIGURATION Config0

	RESOURCE Res0 ON PLC
		TASK task0(INTERVAL := T#20ms,PRIORITY := 0);
		PROGRAM instance0 WITH task0 : program0;
	END_RESOURCE

END_CONFIGURATION

(* ---- 56-DT_TO_TOD.ST ---- *)
FUNCTION DT_TO_TOD2:UDINT
	VAR_INPUT
		IN :	UDINT;
	END_VAR

	DT_TO_TOD2 := (IN MOD UDINT#86400) * UDINT#1000;
END_FUNCTION

PROGRAM program0
  VAR
    LocalVar0 : UDINT;
	LocalOUT  : UDINT;
  END_VAR
  	LocalOUT := DT_TO_TOD2(LocalVar0);
END_PROGRAM

CONFIGURATION Config0
  RESOURCE Res0 ON PLC
    TASK task0(INTERVAL := T#20ms,PRIORITY := 0);
    PROGRAM instance0 WITH task0 : program0;
  END_RESOURCE
END_CONFIGURATION

(* ---- 564-MULTI_IN.ST ---- *)
FUNCTION MID3:REAL

	VAR_INPUT
		IN1 :	REAL;
		IN2 :	REAL;
		IN3 :	REAL;
	END_VAR

	VAR
		_IN1 :	REAL;
		_IN2 :	REAL;
		_IN3 :	REAL;
	END_VAR

	_IN1 := IN1;
	_IN2 := IN2;
	_IN3 := IN3;

	IF _IN1 > _IN2 THEN MID3 := _IN1; _IN1 := _IN2; _IN2 := MID3; END_IF;
	IF _IN2 > _IN3 THEN _IN2 := _IN3; END_IF;
	MID3 := SEL(_IN1 > _IN2, _IN2, _IN1);

END_FUNCTION

FUNCTION _BYTE_TO_INT:INT
	VAR_INPUT
		IN :	BYTE;
	END_VAR

	_BYTE_TO_INT := USINT_TO_INT(BYTE_TO_USINT(IN));
END_FUNCTION

FUNCTION MULTI_IN:REAL

	VAR_INPUT
		IN_1 :	REAL;
		IN_2 :	REAL;
		IN_3 :	REAL;
		DEFAULT :	REAL;
		IN_MIN :	REAL;
		IN_MAX :	REAL;
		MODE :	BYTE;
	END_VAR

	VAR
		count :	INT;
		F1 :	BOOL;
		F2 :	BOOL;
		F3 :	BOOL;
	END_VAR

	F1 :=  in_1 > in_min AND in_1 < in_max;
	F2 :=  in_2 > in_min AND in_2 < in_max;
	F3 :=  in_3 > in_min AND in_3 < in_max;

	CASE _BYTE_TO_INT(mode) OF
	0:	count := 0;
		IF F1 THEN
			count := count + 1;
			MULTI_IN := in_1;
		ELSE
			MULTI_IN := 0.0;
		END_IF;
		IF F2 THEN
			count := count + 1;
			MULTI_IN := MULTI_IN + in_2;
		END_IF;
		IF F3 THEN
			count := count + 1;
			MULTI_IN := MULTI_IN + in_3;
		END_IF;
		MULTI_IN := SEL_REAL(count = 0, MULTI_IN / INT_TO_REAL(count), default);

	1:	MULTI_IN := SEL_REAL(F1, default, IN_1);

	2:	MULTI_IN := SEL_REAL(F2, default, IN_2);

	3:	MULTI_IN := SEL_REAL(F3, default, IN_3);

	4:	MULTI_IN := default;

	5:	MULTI_IN := SEL_REAL(F1, in_max, IN_1);
		IF F2 AND in_2 < MULTI_IN THEN MULTI_IN := in_2; END_IF;
		IF F3 AND in_3 < MULTI_IN THEN MULTI_IN := in_3; END_IF;
		IF MULTI_IN = in_max THEN MULTI_IN := default; END_IF;

	6:	MULTI_IN := SEL_REAL(F1, in_min, IN_1);
		IF F2 AND in_2 > MULTI_IN THEN MULTI_IN := in_2; END_IF;
		IF F3 AND in_3 > MULTI_IN THEN MULTI_IN := in_3; END_IF;
		IF MULTI_IN = in_min THEN MULTI_IN := default; END_IF;

	7:	IF F1 AND F2 AND F3 THEN MULTI_IN := MID3(in_1, in_2, in_3);
		ELSIF F1 AND F2 THEN MULTI_IN := MIN(in_1, in_2);
		ELSIF F1 AND F3 THEN MULTI_IN := MIN(in_1, in_3);
		ELSIF F2 AND F3 THEN MULTI_IN := MIN(in_2, in_3);
		ELSIF F1 THEN MULTI_IN := in_1;
		ELSIF F2 THEN MULTI_IN := in_2;
		ELSIF F3 THEN MULTI_IN := in_3;
		ELSE MULTI_IN := default;
		END_IF;

	END_CASE;

END_FUNCTION

PROGRAM program0
	VAR
		IN_1 :	REAL;
		IN_2 :	REAL;
		IN_3 :	REAL;
		DEFAULT :	REAL;
		IN_MIN :	REAL;
		IN_MAX :	REAL;
		MODE :	BYTE;

		OUT : REAL;
	END_VAR

	OUT := MULTI_IN(IN_1, IN_2, IN_3, DEFAULT, IN_MIN, IN_MAX, MODE);

END_PROGRAM

CONFIGURATION Config0

	RESOURCE Res0 ON PLC
		TASK task0(INTERVAL := T#20ms,PRIORITY := 0);
		PROGRAM instance0 WITH task0 : program0;
	END_RESOURCE

END_CONFIGURATION

(* ---- 567-UTC_TO_LTIME.ST ---- *)
FUNCTION _INT_TO_UDINT:UDINT
	VAR_INPUT
		IN :	INT;
	END_VAR

	_INT_TO_UDINT := DINT_TO_UDINT(INT_TO_DINT(IN));
END_FUNCTION

FUNCTION DT_TO_DATE2:UDINT
	VAR_INPUT
		IN :	UDINT;
	END_VAR

	DT_TO_DATE2 := (IN / UDINT#86400) * UDINT#86400;
END_FUNCTION

FUNCTION YEAR_OF_DATE:INT
	VAR_INPUT
		IDATE :	UDINT;
	END_VAR

	YEAR_OF_DATE := UDINT_TO_INT((idate+UDINT#43200) / UDINT#31557600 + UDINT#1970);
END_FUNCTION

FUNCTION SET_DT:UDINT

	VAR_INPUT
		YEAR : INT;
		MONTH :	INT;
		DAY : INT;
		HOUR : INT;
		MINUTE : INT;
		SECOND : INT;
	END_VAR

	SET_DT := SET_DATE(YEAR, MONTH, DAY) + _INT_TO_UDINT(SECOND) + _INT_TO_UDINT(MINUTE) * UDINT#60 + _INT_TO_UDINT(HOUR) * UDINT#3600;

END_FUNCTION

FUNCTION SET_DATE:UDINT

	VAR_INPUT
		YEAR :	INT;
		MONTH :	INT;
		DAY :	INT;
	END_VAR

	VAR
		count :	INT;
	END_VAR

	IF month > 2 THEN
		count := (month - 1) * 30;
		IF month > 7 THEN
			count := count + DWORD_TO_INT(SHR(DINT_TO_DWORD(INT_TO_DINT(month) - INT_TO_DINT(3)),1));
		ELSE
			count := count + DWORD_TO_INT(SHR(DINT_TO_DWORD(INT_TO_DINT(month) - INT_TO_DINT(4)),1));
		END_IF;
		IF SHL(INT_TO_WORD(year),14) = WORD#0 THEN
			count := count + 1;
		END_IF;
	ELSE
		count := (month - 1) * 31;
	END_IF;
	SET_DATE := (_INT_TO_UDINT(count + day - 1) + DWORD_TO_UDINT(SHR(UDINT_TO_DWORD(_INT_TO_UDINT(year) * UDINT#1461 - UDINT#2878169), 2))) * UDINT#86400;

END_FUNCTION

FUNCTION DST:BOOL
	VAR_INPUT
		UTC :	UDINT;
	END_VAR

	VAR
		yr :	INT;
		yr4 :	UDINT;
		ltc :	UDINT;
		idate :	UDINT;
	END_VAR

	yr := YEAR_OF_DATE(DT_TO_DATE2(UTC));
	ltc := UTC;
	idate := SET_DT(yr, 3, 31, 1, 0, 0);
	yr4 := DWORD_TO_UDINT(SHR(INT_TO_DWORD(5 * yr), 2)) + UDINT#1;
	DST := (idate - ((yr4 + UDINT#3) MOD UDINT#7) * UDINT#86400 <= ltc) AND (idate + (UDINT#214 - (yr4) MOD UDINT#7) * UDINT#86400 > ltc);

END_FUNCTION

FUNCTION UTC_TO_LTIME:UDINT

	VAR_INPUT
		UTC :	UDINT;
		DST_ENABLE :	BOOL;
		TIME_ZONE_OFFSET :	INT;
	END_VAR

	VAR
		tmp :	INT;
	END_VAR

	UTC_TO_LTIME := UTC + _INT_TO_UDINT(TIME_ZONE_OFFSET) * UDINT#60 + BOOL_TO_UDINT(DST_ENABLE AND DST(UTC)) * UDINT#3600;

	tmp := TIME_ZONE_OFFSET * 60 + BOOL_TO_INT(DST_ENABLE AND DST(UTC)) * 3600;
	IF tmp < 0 THEN
		UTC_TO_LTIME := UTC - _INT_TO_UDINT(ABS(tmp));
	ELSE
		UTC_TO_LTIME := UTC + _INT_TO_UDINT(tmp);
	END_IF;

END_FUNCTION

PROGRAM program0
  VAR
	UTC :	UDINT;
	DST_ENABLE :	BOOL;
	TIME_ZONE_OFFSET :	INT;
    CEIL5_OUT : UDINT;
  END_VAR

  CEIL5_OUT := UTC_TO_LTIME(UTC, DST_ENABLE, TIME_ZONE_OFFSET);
END_PROGRAM

CONFIGURATION Config0

  RESOURCE Res0 ON PLC
    TASK task0(INTERVAL := T#20ms,PRIORITY := 0);
    PROGRAM instance0 WITH task0 : program0;
  END_RESOURCE
END_CONFIGURATION

(* ---- 57-MUL_ADD.ST ---- *)
FUNCTION MUL_ADD:REAL

	VAR_INPUT
		X :	REAL;
		K :	REAL;
		O :	REAL;
	END_VAR

	MUL_ADD := X * K + O;

END_FUNCTION

PROGRAM program0
	VAR
		X :	REAL;
		K :	REAL;
		O :	REAL;

		OUT : REAL;
	END_VAR

	OUT := MUL_ADD(X, K, O);

END_PROGRAM

CONFIGURATION Config0

	RESOURCE Res0 ON PLC
		TASK task0(INTERVAL := T#20ms,PRIORITY := 0);
		PROGRAM instance0 WITH task0 : program0;
	END_RESOURCE

END_CONFIGURATION

(* ---- 579-MONTH_END.ST ---- *)
FUNCTION LEAP_OF_DATE:BOOL

	VAR_INPUT
		IDATE :	UDINT;
	END_VAR

	LEAP_OF_DATE := SHL(UDINT_TO_DWORD((idate + UDINT#43200) / UDINT#31557600), 30) = DWORD#16#80000000;
END_FUNCTION

FUNCTION DAY_OF_YEAR:INT
	VAR_INPUT
		IDATE :	UDINT;
	END_VAR

	DAY_OF_YEAR := UDINT_TO_INT(((idate) / UDINT#86400) MOD UDINT#1461);
	IF DAY_OF_YEAR > 729 THEN
		IF DAY_OF_YEAR > 1095 THEN DAY_OF_YEAR := DAY_OF_YEAR - 1095; ELSE DAY_OF_YEAR := DAY_OF_YEAR - 729; END_IF;
	ELSIF DAY_OF_YEAR > 364 THEN
		DAY_OF_YEAR := DAY_OF_YEAR - 364;
	ELSE
		DAY_OF_YEAR := DAY_OF_YEAR + 1;
	END_IF;
END_FUNCTION

FUNCTION MONTH_OF_DATE:INT

	VAR_INPUT
		IDATE :	UDINT;
	END_VAR

	MONTH_OF_DATE := DAY_OF_YEAR(idate);
	IF MONTH_OF_DATE < 32 THEN
		MONTH_OF_DATE := 1;
	ELSIF LEAP_OF_DATE((IDATE)) THEN
		MONTH_OF_DATE := (MONTH_OF_DATE * 53 + 1668) / 1623;
	ELSE
		MONTH_OF_DATE := (MONTH_OF_DATE * 53 + 1700) / 1620;
	END_IF;
END_FUNCTION

FUNCTION YEAR_OF_DATE:INT
	VAR_INPUT
		IDATE :	UDINT;
	END_VAR

	YEAR_OF_DATE := UDINT_TO_INT((idate+UDINT#43200) / UDINT#31557600 + UDINT#1970);
END_FUNCTION

FUNCTION _INT_TO_UDINT:UDINT
	VAR_INPUT
		IN :	INT;
	END_VAR

	_INT_TO_UDINT := DINT_TO_UDINT(INT_TO_DINT(IN));
END_FUNCTION

FUNCTION DT_TO_DATE:UDINT
	VAR_INPUT
		IN :	UDINT;
	END_VAR

	DT_TO_DATE := (IN / UDINT#86400) * UDINT#86400;
END_FUNCTION

FUNCTION SET_DT:UDINT

	VAR_INPUT
		YEAR : INT;
		MONTH :	INT;
		DAY : INT;
		HOUR : INT;
		MINUTE : INT;
		SECOND : INT;
	END_VAR

	SET_DT := SET_DATE(YEAR, MONTH, DAY) + _INT_TO_UDINT(SECOND) + _INT_TO_UDINT(MINUTE) * UDINT#60 + _INT_TO_UDINT(HOUR) * UDINT#3600;

END_FUNCTION

FUNCTION SET_DATE:UDINT

	VAR_INPUT
		YEAR :	INT;
		MONTH :	INT;
		DAY :	INT;
	END_VAR

	VAR
		count :	INT;
	END_VAR

	IF month > 2 THEN
		count := (month - 1) * 30;
		IF month > 7 THEN
			count := count + DWORD_TO_INT(SHR(DINT_TO_DWORD(INT_TO_DINT(month) - INT_TO_DINT(3)),1));
		ELSE
			count := count + DWORD_TO_INT(SHR(DINT_TO_DWORD(INT_TO_DINT(month) - INT_TO_DINT(4)),1));
		END_IF;
		IF SHL(INT_TO_WORD(year),14) = WORD#0 THEN
			count := count + 1;
		END_IF;
	ELSE
		count := (month - 1) * 31;
	END_IF;
	SET_DATE := (_INT_TO_UDINT(count + day - 1) + DWORD_TO_UDINT(SHR(UDINT_TO_DWORD(_INT_TO_UDINT(year) * UDINT#1461 - UDINT#2878169), 2))) * UDINT#86400;

END_FUNCTION

FUNCTION MONTH_END:UDINT

	VAR_INPUT
		IDATE :	UDINT;
	END_VAR

	MONTH_END := SET_DATE(YEAR_OF_DATE(idate),MONTH_OF_DATE(idate)+1,1) - UDINT#86400;

END_FUNCTION

PROGRAM program0
	VAR
		IDATE :	UDINT;

		OUT : UDINT;
	END_VAR

	OUT := MONTH_END(IDATE);

END_PROGRAM

CONFIGURATION Config0

	RESOURCE Res0 ON PLC
		TASK task0(INTERVAL := T#20ms,PRIORITY := 0);
		PROGRAM instance0 WITH task0 : program0;
	END_RESOURCE

END_CONFIGURATION

(* ---- 58-MUX_2.ST ---- *)
FUNCTION MUX_2:BOOL

	VAR_INPUT
		D0 :	BOOL;
		D1 :	BOOL;
		A0 :	BOOL;
	END_VAR

	MUX_2 := SEL(A0, D0, D1);

END_FUNCTION

PROGRAM program0
	VAR
		D0 :	BOOL;
		D1 :	BOOL;
		A0 :	BOOL;
		OUT : BOOL;
	END_VAR

	OUT := MUX_2(D0, D1, A0);

END_PROGRAM

CONFIGURATION Config0

	RESOURCE Res0 ON PLC
		TASK task0(INTERVAL := T#20ms,PRIORITY := 0);
		PROGRAM instance0 WITH task0 : program0;
	END_RESOURCE

END_CONFIGURATION

(* ---- 583-MONTH_BEGIN.ST ---- *)
FUNCTION LEAP_OF_DATE:BOOL

	VAR_INPUT
		IDATE :	UDINT;
	END_VAR

	LEAP_OF_DATE := SHL(UDINT_TO_DWORD((idate + UDINT#43200) / UDINT#31557600), 30) = DWORD#16#80000000;
END_FUNCTION

FUNCTION DAY_OF_YEAR:INT
	VAR_INPUT
		IDATE :	UDINT;
	END_VAR

	DAY_OF_YEAR := UDINT_TO_INT(((idate) / UDINT#86400) MOD UDINT#1461);
	IF DAY_OF_YEAR > 729 THEN
		IF DAY_OF_YEAR > 1095 THEN DAY_OF_YEAR := DAY_OF_YEAR - 1095; ELSE DAY_OF_YEAR := DAY_OF_YEAR - 729; END_IF;
	ELSIF DAY_OF_YEAR > 364 THEN
		DAY_OF_YEAR := DAY_OF_YEAR - 364;
	ELSE
		DAY_OF_YEAR := DAY_OF_YEAR + 1;
	END_IF;
END_FUNCTION

FUNCTION MONTH_OF_DATE:INT

	VAR_INPUT
		IDATE :	UDINT;
	END_VAR

	MONTH_OF_DATE := DAY_OF_YEAR(idate);
	IF MONTH_OF_DATE < 32 THEN
		MONTH_OF_DATE := 1;
	ELSIF LEAP_OF_DATE((IDATE)) THEN
		MONTH_OF_DATE := (MONTH_OF_DATE * 53 + 1668) / 1623;
	ELSE
		MONTH_OF_DATE := (MONTH_OF_DATE * 53 + 1700) / 1620;
	END_IF;
END_FUNCTION

FUNCTION DAY_OF_MONTH:INT
	VAR_INPUT
		IDATE :	UDINT;
	END_VAR

	day_of_month := day_of_year(idate);

	IF leap_of_Date((idate)) THEN
		CASE day_of_month OF
			32..60	:	day_of_month := day_of_month - 31;
			61..91	:	day_of_month := day_of_month - 60;
			92..121 :	day_of_month := day_of_month - 91;
			122..152:	day_of_month := day_of_month - 121;
			153..182:	day_of_month := day_of_month - 152;
			183..213:	day_of_month := day_of_month - 182;
			214..244:	day_of_month := day_of_month - 213;
			245..274:	day_of_month := day_of_month - 244;
			275..305:	day_of_month := day_of_month - 274;
			306..335:	day_of_month := day_of_month - 305;
			336..366:	day_of_month := day_of_month - 335;
		END_CASE;
	ELSE
		CASE day_of_month OF
			32..59	:	day_of_month := day_of_month - 31;
			60..90	:	day_of_month := day_of_month - 59;
			91..120 :	day_of_month := day_of_month - 90;
			121..151:	day_of_month := day_of_month - 120;
			152..181:	day_of_month := day_of_month - 151;
			182..212:	day_of_month := day_of_month - 181;
			213..243:	day_of_month := day_of_month - 212;
			244..273:	day_of_month := day_of_month - 243;
			274..304:	day_of_month := day_of_month - 273;
			305..334:	day_of_month := day_of_month - 304;
			335..365:	day_of_month := day_of_month - 334;
		END_CASE;
	END_IF;
END_FUNCTION

FUNCTION _INT_TO_UDINT:UDINT
	VAR_INPUT
		IN :	INT;
	END_VAR

	_INT_TO_UDINT := DINT_TO_UDINT(INT_TO_DINT(IN));
END_FUNCTION

FUNCTION MONTH_BEGIN:UDINT

VAR_INPUT
	IDATE :	UDINT;
END_VAR

MONTH_BEGIN := idate - _INT_TO_UDINT(DAY_OF_MONTH(idate) - 1) * UDINT#86400;

END_FUNCTION

PROGRAM program0
	VAR
		IDATE :	UDINT;

		OUT : UDINT;
	END_VAR

	OUT := MONTH_BEGIN(IDATE);

END_PROGRAM

CONFIGURATION Config0

	RESOURCE Res0 ON PLC
		TASK task0(INTERVAL := T#20ms,PRIORITY := 0);
		PROGRAM instance0 WITH task0 : program0;
	END_RESOURCE

END_CONFIGURATION

(* ---- 59-_WORD_TO_DINT.ST ---- *)
FUNCTION _WORD_TO_DINT:DINT
	VAR_INPUT
		IN :	WORD;
	END_VAR
	_WORD_TO_DINT := UINT_TO_DINT(WORD_TO_UINT(IN));
END_FUNCTION
PROGRAM program0
  VAR
    LocalVar0 : WORD;
    LocalOUT  : DINT;
  END_VAR

  LocalOUT := _WORD_TO_DINT(LocalVar0);
END_PROGRAM

CONFIGURATION Config0
  RESOURCE Res0 ON PLC
    TASK task0(INTERVAL := T#20ms,PRIORITY := 0);
    PROGRAM instance0 WITH task0 : program0;
  END_RESOURCE
END_CONFIGURATION

(* ---- 6-INV.ST ---- *)
FUNCTION INV:REAL

	VAR_INPUT
		X :	REAL;
	END_VAR

	IF X <> 0.0 THEN INV := 1.0 / X; END_IF;

END_FUNCTION

PROGRAM program0
	VAR
		X :	REAL;
		OUT : REAL;
	END_VAR

	OUT := INV(X);
END_PROGRAM

CONFIGURATION Config0

	RESOURCE Res0 ON PLC
		TASK task0(INTERVAL := T#20ms,PRIORITY := 0);
		PROGRAM instance0 WITH task0 : program0;
	END_RESOURCE

END_CONFIGURATION

(* ---- 60-_BYTE_TO_DINT.ST ---- *)
FUNCTION _BYTE_TO_DINT:DINT
	VAR_INPUT
		IN :	BYTE;
	END_VAR

	_BYTE_TO_DINT := USINT_TO_DINT(BYTE_TO_USINT(IN));
END_FUNCTION

PROGRAM program0
  VAR
    LocalVar0 : BYTE;
	LocalOUT  : DINT;
  END_VAR

  LocalOUT := _BYTE_TO_DINT(LocalVar0);
END_PROGRAM

CONFIGURATION Config0
  RESOURCE Res0 ON PLC
    TASK task0(INTERVAL := T#20ms,PRIORITY := 0);
    PROGRAM instance0 WITH task0 : program0;
  END_RESOURCE
END_CONFIGURATION

(* ---- 61-_BYTE_TO_REAL.ST ---- *)
FUNCTION _BYTE_TO_REAL:REAL
	VAR_INPUT
		IN :	BYTE;
	END_VAR

	_BYTE_TO_REAL := USINT_TO_REAL(BYTE_TO_USINT(IN));
END_FUNCTION

PROGRAM program0
  VAR
    LocalVar0 : BYTE;
	LocalOUT  : REAL;
  END_VAR

  LocalOUT := _BYTE_TO_REAL(LocalVar0);
END_PROGRAM

CONFIGURATION Config0
  RESOURCE Res0 ON PLC
    TASK task0(INTERVAL := T#20ms,PRIORITY := 0);
    PROGRAM instance0 WITH task0 : program0;
  END_RESOURCE
END_CONFIGURATION

(* ---- 62-_INT_TO_UDINT.ST ---- *)
FUNCTION _INT_TO_UDINT:UDINT
	VAR_INPUT
		IN :	INT;
	END_VAR

	_INT_TO_UDINT := DINT_TO_UDINT(INT_TO_DINT(IN));
END_FUNCTION

PROGRAM program0
  VAR
    LocalVar0 : INT;
	LocalOUT  : UDINT;
  END_VAR

  LocalOUT := _INT_TO_UDINT(LocalVar0);
END_PROGRAM

CONFIGURATION Config0
  RESOURCE Res0 ON PLC
    TASK task0(INTERVAL := T#20ms,PRIORITY := 0);
    PROGRAM instance0 WITH task0 : program0;
  END_RESOURCE
END_CONFIGURATION

(* ---- 63-MAX_TIME.ST ---- *)
FUNCTION _MAX_TIME:TIME

	VAR_INPUT
		IN1 :	TIME;
		IN2 :	TIME;
	END_VAR

	_MAX_TIME := SEL_TIME(IN1 < IN2,IN1,IN2);

END_FUNCTION

PROGRAM program0
	VAR
		IN1 :	TIME;
		IN2 :	TIME;

		OUT : TIME;
	END_VAR

	OUT := _MAX_TIME(IN1, IN2);

END_PROGRAM

CONFIGURATION Config0

	RESOURCE Res0 ON PLC
		TASK task0(INTERVAL := T#20ms,PRIORITY := 0);
		PROGRAM instance0 WITH task0 : program0;
	END_RESOURCE

END_CONFIGURATION

(* ---- 64-SECOND_OF_DT.ST ---- *)
FUNCTION SECOND_OF_DT:INT

	VAR_INPUT
		XDT :	UDINT;
	END_VAR

	SECOND_OF_DT := UDINT_TO_INT(XDT MOD UDINT#60);
END_FUNCTION

PROGRAM program0
  VAR
    LocalVar0 : UDINT;
	LocalOUT  : INT;
  END_VAR
  	LocalOUT := SECOND_OF_DT(LocalVar0);
END_PROGRAM

CONFIGURATION Config0
  RESOURCE Res0 ON PLC
    TASK task0(INTERVAL := T#20ms,PRIORITY := 0);
    PROGRAM instance0 WITH task0 : program0;
  END_RESOURCE
END_CONFIGURATION

(* ---- 65-UDINT_TO_TIME.ST ---- *)
FUNCTION _UDINT_TO_TIME:TIME

	VAR_INPUT
		IN :	UDINT;
	END_VAR

	_UDINT_TO_TIME := DINT_TO_TIME(UDINT_TO_DINT(IN));

END_FUNCTION

PROGRAM program0
  VAR
	  IN :	UDINT;
    CEIL5_OUT : TIME;
  END_VAR

  CEIL5_OUT := _UDINT_TO_TIME(IN);
END_PROGRAM

CONFIGURATION Config0

  RESOURCE Res0 ON PLC
    TASK task0(INTERVAL := T#20ms,PRIORITY := 0);
    PROGRAM instance0 WITH task0 : program0;
  END_RESOURCE
END_CONFIGURATION

(* ---- 66-_WORD_TO_REAL.ST ---- *)
FUNCTION _WORD_TO_REAL:REAL
	VAR_INPUT
		IN :	WORD;
	END_VAR
	_WORD_TO_REAL := UINT_TO_REAL(WORD_TO_UINT(IN));
END_FUNCTION

PROGRAM program0
  VAR
    LocalVar0 : WORD;
    LocalOUT  : REAL;
  END_VAR

  LocalOUT := _WORD_TO_REAL(LocalVar0);
END_PROGRAM

CONFIGURATION Config0
  RESOURCE Res0 ON PLC
    TASK task0(INTERVAL := T#20ms,PRIORITY := 0);
    PROGRAM instance0 WITH task0 : program0;
  END_RESOURCE
END_CONFIGURATION

(* ---- 662-DATE_ADD.ST ---- *)
FUNCTION YEAR_OF_DATE:INT
	VAR_INPUT
		IDATE :	UDINT;
	END_VAR

	YEAR_OF_DATE := UDINT_TO_INT((idate+UDINT#43200) / UDINT#31557600 + UDINT#1970);
END_FUNCTION

FUNCTION DAY_OF_WEEK:INT

	VAR_INPUT
		IDATE :	UDINT;
	END_VAR

	DAY_OF_WEEK := UDINT_TO_INT((idate / UDINT#86400 + UDINT#3) MOD UDINT#7) + INT#01;
END_FUNCTION

FUNCTION LEAP_OF_DATE:BOOL

	VAR_INPUT
		IDATE :	UDINT;
	END_VAR

	LEAP_OF_DATE := SHL(UDINT_TO_DWORD((idate + UDINT#43200) / UDINT#31557600), 30) = DWORD#16#80000000;
END_FUNCTION

FUNCTION DAY_OF_YEAR:INT
	VAR_INPUT
		IDATE :	UDINT;
	END_VAR

	DAY_OF_YEAR := UDINT_TO_INT(((idate) / UDINT#86400) MOD UDINT#1461);
	IF DAY_OF_YEAR > 729 THEN
		IF DAY_OF_YEAR > 1095 THEN DAY_OF_YEAR := DAY_OF_YEAR - 1095; ELSE DAY_OF_YEAR := DAY_OF_YEAR - 729; END_IF;
	ELSIF DAY_OF_YEAR > 364 THEN
		DAY_OF_YEAR := DAY_OF_YEAR - 364;
	ELSE
		DAY_OF_YEAR := DAY_OF_YEAR + 1;
	END_IF;
END_FUNCTION

FUNCTION MONTH_OF_DATE:INT

	VAR_INPUT
		IDATE :	UDINT;
	END_VAR

	MONTH_OF_DATE := DAY_OF_YEAR(idate);
	IF MONTH_OF_DATE < 32 THEN
		MONTH_OF_DATE := 1;
	ELSIF LEAP_OF_DATE((IDATE)) THEN
		MONTH_OF_DATE := (MONTH_OF_DATE * 53 + 1668) / 1623;
	ELSE
		MONTH_OF_DATE := (MONTH_OF_DATE * 53 + 1700) / 1620;
	END_IF;
END_FUNCTION

FUNCTION DAY_OF_MONTH:INT
	VAR_INPUT
		IDATE :	UDINT;
	END_VAR

	day_of_month := day_of_year(idate);

	IF leap_of_Date((idate)) THEN
		CASE day_of_month OF
			32..60	:	day_of_month := day_of_month - 31;
			61..91	:	day_of_month := day_of_month - 60;
			92..121 :	day_of_month := day_of_month - 91;
			122..152:	day_of_month := day_of_month - 121;
			153..182:	day_of_month := day_of_month - 152;
			183..213:	day_of_month := day_of_month - 182;
			214..244:	day_of_month := day_of_month - 213;
			245..274:	day_of_month := day_of_month - 244;
			275..305:	day_of_month := day_of_month - 274;
			306..335:	day_of_month := day_of_month - 305;
			336..366:	day_of_month := day_of_month - 335;
		END_CASE;
	ELSE
		CASE day_of_month OF
			32..59	:	day_of_month := day_of_month - 31;
			60..90	:	day_of_month := day_of_month - 59;
			91..120 :	day_of_month := day_of_month - 90;
			121..151:	day_of_month := day_of_month - 120;
			152..181:	day_of_month := day_of_month - 151;
			182..212:	day_of_month := day_of_month - 181;
			213..243:	day_of_month := day_of_month - 212;
			244..273:	day_of_month := day_of_month - 243;
			274..304:	day_of_month := day_of_month - 273;
			305..334:	day_of_month := day_of_month - 304;
			335..365:	day_of_month := day_of_month - 334;
		END_CASE;
	END_IF;
END_FUNCTION

FUNCTION _INT_TO_UDINT:UDINT
	VAR_INPUT
		IN :	INT;
	END_VAR

	_INT_TO_UDINT := DINT_TO_UDINT(INT_TO_DINT(IN));
END_FUNCTION

FUNCTION SET_DATE:UDINT

	VAR_INPUT
		YEAR :	INT;
		MONTH :	INT;
		DAY :	INT;
	END_VAR

	VAR
		count :	INT;
	END_VAR

	IF month > 2 THEN
		count := (month - 1) * 30;
		IF month > 7 THEN
			count := count + DWORD_TO_INT(SHR(DINT_TO_DWORD(INT_TO_DINT(month) - INT_TO_DINT(3)),1));
		ELSE
			count := count + DWORD_TO_INT(SHR(DINT_TO_DWORD(INT_TO_DINT(month) - INT_TO_DINT(4)),1));
		END_IF;
		IF SHL(INT_TO_WORD(year),14) = WORD#0 THEN
			count := count + 1;
		END_IF;
	ELSE
		count := (month - 1) * 31;
	END_IF;
	SET_DATE := (_INT_TO_UDINT(count + day - 1) + DWORD_TO_UDINT(SHR(UDINT_TO_DWORD(_INT_TO_UDINT(year) * UDINT#1461 - UDINT#2878169), 2))) * UDINT#86400;

END_FUNCTION

FUNCTION DATE_ADD:UDINT
	VAR_INPUT
		IDATE :	UDINT;
		D :	INT;
		W :	INT;
		M :	INT;
		Y :	INT;
	END_VAR

	VAR
		mo :	INT;
		yr :	INT;
		dm :	INT;
	END_VAR

	DATE_ADD := IDATE + INT_TO_UDINT(D + W * 7) * UDINT#86400;
	yr := Y + YEAR_OF_DATE(DATE_ADD);
	mo := M + MONTH_OF_DATE(DATE_ADD);
	dm := DAY_OF_MONTH(DATE_ADD);
	WHILE mo > 12 DO
		mo := mo - 12;
		yr := yr + 1;
	END_WHILE;
	WHILE mo < 1 DO
		mo := mo + 12;
		yr := yr - 1;
	END_WHILE;
	DATE_ADD := SET_DATE(yr, mo, dm);
END_FUNCTION

PROGRAM program0
  VAR
    LocalVar0 : UDINT;
	LocalVar1 : INT;
	LocalVar2 : INT;
	LocalVar3 : INT;
	LocalVar4 : INT;
	LocalOUT  : UDINT;
  END_VAR
  	LocalOUT := DATE_ADD(LocalVar0, LocalVar1, LocalVar2, LocalVar3, LocalVar4);
END_PROGRAM

CONFIGURATION Config0
  RESOURCE Res0 ON PLC
    TASK task0(INTERVAL := T#20ms,PRIORITY := 0);
    PROGRAM instance0 WITH task0 : program0;
  END_RESOURCE
END_CONFIGURATION

(* ---- 67-TIME_TO_DWORD.ST ---- *)
FUNCTION TIME_TO_DWORD1:DWORD

VAR_INPUT
	X :	TIME;
END_VAR

TIME_TO_DWORD1 := UDINT_TO_DWORD(DINT_TO_UDINT(TIME_TO_DINT(X)));
END_FUNCTION

PROGRAM program0
  VAR
	X :	TIME;
    CEIL5_OUT : DWORD;
  END_VAR

  CEIL5_OUT := TIME_TO_DWORD1(X);
END_PROGRAM

CONFIGURATION Config0

  RESOURCE Res0 ON PLC
    TASK task0(INTERVAL := T#20ms,PRIORITY := 0);
    PROGRAM instance0 WITH task0 : program0;
  END_RESOURCE
END_CONFIGURATION

(* ---- 68-DAY_OF_DATE.ST ---- *)
FUNCTION DAY_OF_DATE:DINT
	VAR_INPUT
		IDATE :	UDINT;
	END_VAR

	day_of_date := UDINT_TO_DINT(idate / UDINT#86400);
END_FUNCTION

PROGRAM program0
  VAR
    LocalVar0 : UDINT;
	LocalOUT  : DINT;
  END_VAR
  	LocalOUT := DAY_OF_DATE(LocalVar0);
END_PROGRAM

CONFIGURATION Config0
  RESOURCE Res0 ON PLC
    TASK task0(INTERVAL := T#20ms,PRIORITY := 0);
    PROGRAM instance0 WITH task0 : program0;
  END_RESOURCE
END_CONFIGURATION

(* ---- 69-DWORD_TO_TIME.ST ---- *)
FUNCTION DWORD_TO_TIME2:TIME
	VAR_INPUT
		X :	DWORD;
	END_VAR
	DWORD_TO_TIME2 := DINT_TO_TIME(DWORD_TO_DINT(X));
END_FUNCTION

PROGRAM program0
  VAR
    LocalVar0 : DWORD;
	  LocalOUT  : TIME;
  END_VAR
  	LocalOUT := DWORD_TO_TIME2(LocalVar0);
END_PROGRAM

CONFIGURATION Config0
  RESOURCE Res0 ON PLC
    TASK task0(INTERVAL := T#20ms,PRIORITY := 0);
    PROGRAM instance0 WITH task0 : program0;
  END_RESOURCE
END_CONFIGURATION

(* ---- 7-MS_TO_KMH.ST ---- *)
FUNCTION MS_TO_KMH:REAL

	VAR_INPUT
		MS :	REAL;
	END_VAR

	MS_TO_KMH := Ms * 3.6;

END_FUNCTION

PROGRAM program0
	VAR
		MS :	REAL;

		OUT : REAL;
	END_VAR

	OUT := MS_TO_KMH(MS);

END_PROGRAM

CONFIGURATION Config0

	RESOURCE Res0 ON PLC
		TASK task0(INTERVAL := T#20ms,PRIORITY := 0);
		PROGRAM instance0 WITH task0 : program0;
	END_RESOURCE

END_CONFIGURATION

(* ---- 70-SHL1.ST ---- *)
FUNCTION SHL1:DWORD

	VAR_INPUT
		IN :	DWORD;
		N :	INT;
	END_VAR

	SHL1 := SHR(DWORD#16#FF_FF_FF_FF,32-N) OR SHL(IN,N);

END_FUNCTION

PROGRAM program0

	VAR
		IN :	DWORD;
		N :	INT;
		CEIL5_OUT : DWORD;
	END_VAR

  	CEIL5_OUT := SHL1(IN, N);

END_PROGRAM

CONFIGURATION Config0

	RESOURCE Res0 ON PLC
		TASK task0(INTERVAL := T#20ms,PRIORITY := 0);
		PROGRAM instance0 WITH task0 : program0;
	END_RESOURCE

END_CONFIGURATION

(* ---- 71-SHR1.ST ---- *)
FUNCTION SHR1:DWORD

	VAR_INPUT
		IN :	DWORD;
		N :	INT;
	END_VAR

	SHR1 := SHL(DWORD#16#FF_FF_FF_FF,32-N) OR SHR(IN,N);

END_FUNCTION

PROGRAM program0

	VAR
		IN : DWORD;
		N :	INT;
		CEIL5_OUT : DWORD;
	END_VAR

	CEIL5_OUT := SHR1(IN, N);

END_PROGRAM

CONFIGURATION Config0

	RESOURCE Res0 ON PLC
		TASK task0(INTERVAL := T#20ms,PRIORITY := 0);
		PROGRAM instance0 WITH task0 : program0;
	END_RESOURCE

END_CONFIGURATION

(* ---- 72-INC1.ST ---- *)
FUNCTION INC1:INT

	VAR_INPUT
		X :	INT;
		N :	INT;
	END_VAR

	IF X >= N - 1 THEN
		INC1 := 0;
	ELSE
		INC1 := X + 1;
	END_IF;
END_FUNCTION

PROGRAM program0
  VAR
	X :	INT;
	N :	INT;
    CEIL5_OUT : INT;
  END_VAR

  CEIL5_OUT := INC1(X, N);
END_PROGRAM

CONFIGURATION Config0

  RESOURCE Res0 ON PLC
    TASK task0(INTERVAL := T#20ms,PRIORITY := 0);
    PROGRAM instance0 WITH task0 : program0;
  END_RESOURCE
END_CONFIGURATION

(* ---- 73-_DWORD_TO_REAL.ST ---- *)
FUNCTION _DWORD_TO_REAL:REAL
	VAR_INPUT
		IN :	DWORD;
	END_VAR

	_DWORD_TO_REAL := UDINT_TO_REAL(DWORD_TO_UDINT(IN));
END_FUNCTION

PROGRAM program0
  VAR
    LocalVar0 : DWORD;
    LocalOUT  : REAL;
  END_VAR

  LocalOUT := _DWORD_TO_REAL(LocalVar0);
END_PROGRAM

CONFIGURATION Config0
  RESOURCE Res0 ON PLC
    TASK task0(INTERVAL := T#20ms,PRIORITY := 0);
    PROGRAM instance0 WITH task0 : program0;
  END_RESOURCE
END_CONFIGURATION

(* ---- 74-MUX_R2.ST ---- *)
FUNCTION MUX_R2:REAL

	VAR_INPUT
		IN0 :	REAL;
		IN1 :	REAL;
		A :	BOOL;
	END_VAR

	MUX_R2 := SEL(A, IN0, IN1);

END_FUNCTION

PROGRAM program0
	VAR
		IN0 :	REAL;
		IN1 :	REAL;
		A :	BOOL;

		OUT : REAL;
	END_VAR

	OUT := MUX_R2(IN0, IN1, A);

END_PROGRAM

CONFIGURATION Config0

	RESOURCE Res0 ON PLC
		TASK task0(INTERVAL := T#20ms,PRIORITY := 0);
		PROGRAM instance0 WITH task0 : program0;
	END_RESOURCE

END_CONFIGURATION
